Universal Robots PolyScope program: AdientTorsF_Eol1L.urp

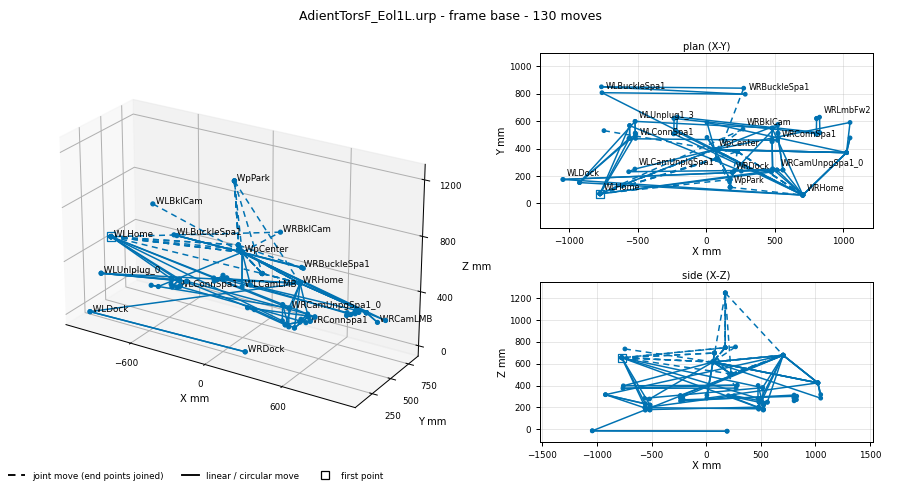
[picture p0: tool path of AdientTorsF_Eol1L.urp in frame base, 130 of 170 moves have a stored position in this frame; points joined in program order, loops and branches not executed]
Program AdientTorsF_Eol1L (installation=EOL_1L directory=/programs createdIn=3.5.1 lastSavedIn=5.26.0 robotSerialNumber=20265101875)
Calibrated DH parameters: a=[-0.000091, -0.609283, -0.566309, 0.000078, -0.000019, 0]; d=[0.180883, 55.684211, -64.380909, 8.871165, 0.119736, 0.115499]; alpha=[1.570556, -0.001038, 0.008646, 1.570192, -1.569654, 0]; deltaTheta=[0, -0.094548, 6.245733, 0.132006, -0.000002, 0]
InitVariablesNode variables(variable(name=Abort, expression=False), variable(name=AdapterReady_L, expression=False), variable(name=AdapterReady_R, expression=False), variable(name=CMD_Heartbt_i1, expression=0), variable(name=CMD_Heartbt_i2, expression=0), variable(name=CMD_Program_i1, expression=0), variable(name=CMD_Program_i2, expression=0), variable(name=CMD_Reserve_i1, expression=0), variable(name=CMD_Reserve_i2, expression=0), variable(name=CMD_Timeout_i1, expression=0), variable(name=CMD_Timeout_i2, expression=0), variable(name=CamCorrectnOK, expression=0), variable(name=DEBUG, expression=False), variable(name=D_rel, expression=p[0,0,0,0,0,0]), variable(name=EvtBeep, expression=False), variable(name=EvtDock, expression=0), variable(name=Mute, expression=False), variable(name=P_ini, expression=get_actual_tcp_pose()), variable(name=Parking, expression=0), variable(name=ProgExe, expression=0), variable(name=STS_Heartbeat, expression=False), variable(name=STS_Progress, expression=0), variable(name=STS_Reservation, expression=0), variable(name=SetCameraProg, expression=0))
BeforeStart
  SuppressedNode
    DEBUG := True
  'SW version, to be used to track changes and keep sync of all stations'
  SW_Ver := 1.0
  Folder Scripts [hidden by the author, left out]
  Folder Avoid guidance screen [hidden by the author, left out]
  Call GripperOpen
  GoToHome := True
  Script: socket_open("127.0.0.1",30001)
Robot Program (runOnlyOnce=false)
  Folder Execute Program
    Folder Init
      Wait Condition expression=EvtDock≤0
      Folder Verify adapter ready
        If digital_in[0] or analog_in[3]<(ivGripSensOpen+0.3)
          AdapterReady_L := False
        If digital_in[4] or analog_in[3]<(ivGripSensOpen+0.3)
          AdapterReady_R := False
      Folder Go to home pos automatically
        If GoToHome and  not (AdapterReady_L or AdapterReady_R)
          Wait Sleep waitTime=1
          If InRange(P_Flange[0],-1,-0.2) and InRange(P_Flange[1],-0.5,0.5) and InRange(P_Flange[2],0.3,1)
            If AdapterDocked or DEBUG or (analog_in[3]<(ivGripSensOpen+0.3))
              MoveJ speed 120 deg/s, acceleration 500 deg/s^2 (useActiveTCP=false positionType=JointAngles optimoveEnabled=false optiMoveSpeed=0.3 optiMoveAcceleration=0.09) tcp=t0_Flange; feature=Base
                Waypoint WLHome: TCP in base x=-773.534 y=70.689 z=655.308 mm, rx=3.1416 ry=0 rz=0 rad; joints [187.663, -96.209, -85.791, -88.066, 90.49, -82.232] deg; TCP offset x=0 y=0 z=0 mm, rx=0 ry=0 rz=3.1416 rad
            Else 
              Popup Error (haltProgram=false message=Adapter must be docked inputType=Text)
              Halt
          ElseIf AtCenterPos
            MoveJ speed 120 deg/s, acceleration 500 deg/s^2 (useActiveTCP=true positionType=JointAngles optimoveEnabled=false optiMoveSpeed=0.3 optiMoveAcceleration=0.09) feature=Base
              Waypoint WpCenter: TCP in base x=62.197 y=393.251 z=616.502 mm, rx=-0.0356 ry=3.1413 rz=-0.0001 rad; joints [106.827, -57.183, -119.283, -93.604, 90.531, 15.582] deg
          ElseIf AtParkPos
            MoveJ speed 120 deg/s, acceleration 500 deg/s^2 (useActiveTCP=true positionType=JointAngles optimoveEnabled=false optiMoveSpeed=0.3 optiMoveAcceleration=0.09) feature=Base
              Waypoint WpPark: TCP in base x=175.046 y=118.455 z=1248.983 mm, rx=-2.2111 ry=2.2293 rz=-0.0002 rad; joints [89.999, -90, 0, -180, 90, -90] deg
          ElseIf InRange(P_Flange[0],0.2,1.2) and InRange(P_Flange[1],-0.5,0.5) and InRange(P_Flange[2],0.3,1)
            If AdapterDocked or DEBUG or (analog_in[3]<(ivGripSensOpen+0.3))
              MoveJ speed 120 deg/s, acceleration 500 deg/s^2 (useActiveTCP=true positionType=JointAngles optimoveEnabled=false optiMoveSpeed=0.3 optiMoveAcceleration=0.09) feature=Base
                Waypoint WRHome: TCP in base x=704.968 y=61.356 z=678.212 mm, rx=-2.2214 ry=-2.2214 rz=0 rad; joints [19.143, -89.513, -90.55, -90.002, 90.503, 19.233] deg; TCP offset x=0 y=0 z=0 mm, rx=0 ry=0 rz=3.1416 rad
            Else 
              Popup Error (haltProgram=false message=Adapter must be docked inputType=Text)
              Halt
          Else 
            Popup Error (haltProgram=false message=Illegal position. Adjust arm to open space in front of the backrest, or [Move]->[Home] inputType=Text)
            Halt
        GoToHome := False
      If DEBUG
        'Popup window with program selection'
        ProgExe :=  (valueSource=Operator message=Program number? valueType=Integer)
      If ProgExe>0
        Folder Init
          Mute := False
          Wait Condition expression=not GoToHome
          If In(ProgExe,[11,12,14])
            AdapterReady_R := False
          ElseIf In(ProgExe,[51,52,54])
            AdapterReady_L := False
          Else 
            AdapterReady_L := False
            AdapterReady_R := False
    Folder Programs
      If InRange(ProgExe,1,99)
        Folder Undock
          If In(ProgExe,[11,51])
            Script: Report(1)
            Folder AtHome?
              Timer (action=Reset) variable(name=T_Timeout)
              Timer (action=Start) variable=T_Timeout
              Wait Condition expression=AtHomePos or T_Timeout>5
              If not AtHomePos
                Script: Report(90)
            If Progress_run() and  not AdapterDocked
              Script: Report(94)
            If Progress_run()
              Folder Undock
                MoveL speed 1000 mm/s, acceleration 3000 mm/s^2 (useActiveTCP=false optimoveEnabled=false optiMoveSpeed=0.3 optiMoveAcceleration=0.09) tcp=t2_Gripper; feature=Base
                  Call GripperOpenQuick
                  If False
                    Waypoint WLDock: TCP in base x=-1043.478 y=175.197 z=-14.02 mm, rx=1.8607 ry=1.8607 rz=0.6057 rad; joints [179.892, -126.837, -85.911, -93.381, 90.434, -0.034] deg; TCP offset x=0 y=-260 z=74 mm, rx=0 ry=0 rz=0 rad
                    Waypoint WRDock: TCP in base x=191.182 y=225.632 z=-17.704 mm, rx=1.8937 ry=1.8608 rz=0.5985 rad; joints [64.532, -92.299, -158.794, -2.395, 58.985, 241.468] deg
                  If ProgExe<50
                    WpDock := WLDock
                    WpHome := WLHome
                  Else 
                    WpDock := WRDock
                    WpHome := WRHome
                  Wp := pose_trans(WpDock, p[0,0.175,-0.1,0,0,0])
                  Waypoint Variable (Variable): motionParameters(blendRadius=0.05); variable=Wp
                  Call GripperOpen
                  Wp := pose_trans(WpDock, p[0,0.075,0.01,0,0,0])
                  Waypoint Variable (Variable): motionParameters(blendRadius=0.01); variable=Wp
                  Wp := pose_trans(WpDock, p[0,0.055,0,0,0,0])
                  Waypoint Variable (Variable): motionParameters(blendRadius=0.01); variable=Wp
                  Waypoint Variable (Variable): variable=WpDock
                  Call GripperClose
                  Wp := pose_trans(WpDock, p[0,0.25,0,0,0,0])
                  Waypoint Variable (Variable): variable=Wp
                If ProgExe<50
                  AdapterReady_L := True
                Else 
                  AdapterReady_R := True
                Script: Report(50)
            Script: Report(50)
        Folder Connect
          If In(ProgExe,[12,14,52,54])
            Script: Report(1)
            If ProgExe<50 and AdapterReady_L
              Undock := False
            ElseIf ProgExe≥50 and AdapterReady_R
              Undock := False
            Else 
              Undock := True
              Folder AtHome? [hidden by the author, left out]
              If Progress_run() and  not AdapterDocked
                Script: Report(94)
            If Progress_run()
              Folder Undock
                If Undock
                  MoveL speed 1000 mm/s, acceleration 3000 mm/s^2 (useActiveTCP=false optimoveEnabled=false optiMoveSpeed=0.3 optiMoveAcceleration=0.09) tcp=t2_Gripper; feature=Base
                    Call GripperOpenQuick
                    If False
                      Waypoint WLDock: TCP in base x=-1043.478 y=175.197 z=-14.02 mm, rx=1.8607 ry=1.8607 rz=0.6057 rad; joints [179.892, -126.837, -85.911, -93.381, 90.434, -0.034] deg; TCP offset x=0 y=-260 z=74 mm, rx=0 ry=0 rz=0 rad
                      Waypoint WRDock: TCP in base x=191.182 y=225.632 z=-17.704 mm, rx=1.8937 ry=1.8608 rz=0.5985 rad; joints [64.532, -92.299, -158.794, -2.395, 58.985, 241.468] deg
                    If ProgExe<50
                      WpDock := WLDock
                      WpHome := WLHome
                    Else 
                      WpDock := WRDock
                      WpHome := WRHome
                    Wp := pose_trans(WpDock, p[0,0.175,-0.1,0,0,0])
                    Waypoint Variable (Variable): motionParameters(blendRadius=0.05); variable=Wp
                    Call GripperOpen
                    Wp := pose_trans(WpDock, p[0,0.075,0.01,0,0,0])
                    Waypoint Variable (Variable): motionParameters(blendRadius=0.01); variable=Wp
                    Wp := pose_trans(WpDock, p[0,0.055,0,0,0,0])
                    Waypoint Variable (Variable): motionParameters(blendRadius=0.01); variable=Wp
                    Waypoint Variable (Variable): variable=WpDock
                    Call GripperClose
                    Wp := pose_trans(WpDock, p[0,0.25,0,0,0,0])
                    Waypoint Variable (Variable): variable=Wp
                AdapterReady_L := False
                AdapterReady_R := False
                Script: Report(2)
              CamCorrection := p[0,0,0,0,0,0]
              SuppressedNode
                Folder Camera
                  MoveL speed 250 mm/s, acceleration 1200 mm/s^2 (useActiveTCP=false optimoveEnabled=false optiMoveSpeed=0.3 optiMoveAcceleration=0.09) tcp=t0_Flange; feature=Base
                    If In(ProgExe,[12,13])
                      SetCameraProg := 12
                      Waypoint WLCamConSpa1: TCP in base x=-511.083 y=256.44 z=253.227 mm, rx=2.1948 ry=2.1949 rz=-0.0574 rad; joints [170.312, -93.988, -133.728, -42.837, 93.248, -9.279] deg; TCP offset x=0 y=0 z=0 mm, rx=0 ry=0 rz=0 rad
                    If In(ProgExe,[14])
                      SetCameraProg := ProgExe
                      Waypoint WLCamConSpa3: TCP in base x=-559.049 y=229.366 z=263.196 mm, rx=-2.2214 ry=-2.2215 rz=0 rad; joints [174.302, -95.829, -130.307, -43.928, 90.296, -5.276] deg
                    If In(ProgExe,[52,53])
                      SetCameraProg := 52
                      Waypoint WRCamConSpa1: TCP in base x=528.577 y=256.538 z=254.589 mm, rx=2.1946 ry=2.1948 rz=-0.0575 rad; joints [43.439, -94.974, -131.929, -45.242, 88.117, 223.892] deg
                    If In(ProgExe,[54])
                      SetCameraProg := ProgExe
                      Waypoint WRCamConSpa3: TCP in base x=480.455 y=221.374 z=266.967 mm, rx=-2.2214 ry=-2.2215 rz=-0.0001 rad; joints [43.801, -88.335, -137.68, -44.047, 90.305, 224.222] deg
                  Call CamAcquire
                  CamCorrection := p[CamData[0],CamData[1]*-0.5,CamData[1],0,0,0]
            SuppressedNode
              If Progress_run() and CamCorrectnOK≠ProgExe
                EvtDock := 1
                Wait Condition expression=EvtDock≟0
                Script: Report(91)
            Folder Connect
              If Progress_run()
                Set NoAction tcp=t2_Gripper
                MoveL speed 1000 mm/s, acceleration 3000 mm/s^2 (useActiveTCP=false optimoveEnabled=false optiMoveSpeed=0.3 optiMoveAcceleration=0.09) tcp=t2_Gripper; feature=Base
                  If False
                    'wp is set to position exactly 30mm below'
                    Waypoint WLConnSpa1: motionParameters(blendRadius=0.045); TCP in base x=-514.347 y=474.559 z=185.987 mm, rx=3.0892 ry=0 rz=0.0001 rad; joints [174.313, -90.885, -134.162, -45.296, 93.296, -95.282] deg; TCP offset x=0 y=260 z=74 mm, rx=0 ry=0 rz=3.1416 rad
                    Waypoint WLConnSpa3: TCP in base x=-563.167 y=472.162 z=197.967 mm, rx=2.9544 ry=0 rz=0.0002 rad; joints [172.16, -92.445, -126.338, -52.702, 100.982, -97.611] deg
                    Waypoint WRConnSpa1: TCP in base x=520.916 y=460.286 z=187.058 mm, rx=3.089 ry=0 rz=-0.0005 rad; joints [39.919, -90.524, -133.875, -47.63, 88.028, 130.365] deg
                    Waypoint WRConnSpa3: TCP in base x=478.559 y=467.416 z=198.199 mm, rx=3.0125 ry=0.0525 rz=-0.0035 rad; joints [44.279, -85.291, -133.969, -56.002, 85.12, 132.879] deg
                  If In(ProgExe,[12])
                    Wp := pose_trans(WLConnSpa1, CamCorrection)
                  If In(ProgExe,[14])
                    Wp := pose_add(WLConnSpa3, CamCorrection)
                  If In(ProgExe,[52])
                    Wp := pose_trans(WRConnSpa1, CamCorrection)
                  If In(ProgExe,[54])
                    Wp := pose_add(WRConnSpa3, CamCorrection)
                  Waypoint Variable (Variable): variable=Wp
                Force Frame feature=Joint_6_name; selection=[0, 0, 1, 0, 0, 0]; wrench=[0, 0, -30, 0, 0, 0]; limitsForce=[0.15, 0.15, 0.1, 1.047198, 1.047198, 1.047198]; limitsMotion=[0.1, 0.1, 0.1, 0.349066, 0.349066, 0.349066]
                  Wait Sleep waitTime=1
                Force Frame feature=Joint_6_name; selection=[1, 0, 1, 0, 0, 0]; wrench=[0, 0, -30, 0, 0, 0]; limitsForce=[0.15, 0.15, 0.05, 1.047198, 1.047198, 1.047198]; limitsMotion=[0.1, 0.1, 0.1, 0.349066, 0.349066, 0.349066]
                  Wait Sleep waitTime=0.5
                'position ok'
                If InRange(Wp[2]+0.03-P_act[2],-0.015,0.015)
                  'ok'
                Else 
                  EvtDock := 2
                  Wait Condition expression=EvtDock≤0
                  Script: Report(96)
              If Progress_run()
                Force Frame feature=Joint_6_name; selection=[0, 1, 0, 0, 0, 0]; wrench=[0, -60, -10, 0, 0, 0]; limitsForce=[0.15, 0.05, 0.01, 1.047198, 1.047198, 1.047198]; limitsMotion=[0.1, 0.1, 0.1, 0.349066, 0.349066, 0.349066]
                  Wait Sleep waitTime=1
                MoveL speed 1000 mm/s, acceleration 3000 mm/s^2 (useActiveTCP=true optimoveEnabled=false optiMoveSpeed=0.3 optiMoveAcceleration=0.09) feature=Base
                  Wp := pose_trans(P_act, p[0,0.005,0,0,0,0])
                  Waypoint Variable (Variable): variable=Wp
                Call GripperOpen
                Force Frame feature=Joint_6_name; selection=[0, 1, 0, 0, 0, 0]; wrench=[0, -60, -10, 0, 0, 0]; limitsForce=[0.15, 0.1, 0.01, 1.047198, 1.047198, 1.047198]; limitsMotion=[0.1, 0.1, 0.1, 0.349066, 0.349066, 0.349066]
                  Wait Sleep waitTime=1
                  Script: Report(5)
                  MoveL speed 500 mm/s, acceleration 2000 mm/s^2 (useActiveTCP=true optimoveEnabled=false optiMoveSpeed=0.3 optiMoveAcceleration=0.09) feature=Base
                    Wp0 := get_actual_tcp_pose()
                    Wp := pose_trans(Wp0, p[0,0,0,0,0,0.07])
                    Waypoint Variable (Variable): variable=Wp
                    Wp := pose_trans(Wp0, p[0,0,0,0,0,-0.07])
                    Waypoint Variable (Variable): variable=Wp
                    Waypoint Variable (Variable): variable=Wp0
                    Wp := pose_trans(Wp0, p[0,0,0.01,0,0,0])
                    Waypoint Variable (Variable): variable=Wp
                    Waypoint Variable (Variable): variable=Wp0
                MoveL speed 1000 mm/s, acceleration 3000 mm/s^2 (useActiveTCP=true optimoveEnabled=false optiMoveSpeed=0.3 optiMoveAcceleration=0.09) feature=Base
                  Wp0 := get_actual_tcp_pose()
                  Wp := pose_trans(Wp0, p[0,0.015,0,0,0,0])
                  Waypoint Variable (Variable): variable=Wp
                Force Frame feature=Joint_6_name; selection=[0, 1, 0, 0, 0, 0]; wrench=[0, -60, 0, 0, 0, 0]; limitsForce=[0.15, 0.5, 0.15, 1.047198, 1.047198, 1.047198]; limitsMotion=[0.1, 0.1, 0.1, 0.349066, 0.349066, 0.349066]
                  Wait Sleep waitTime=0.5
                Script: Report(6)
                Timer (action=Reset) variable=T_Timeout
                Timer (action=Start) variable=T_Timeout
                Folder Test switch pin, retreat on fail
                  Wait Condition expression=Flags[0] or T_Timeout>10 or DEBUG
                  If not Flags[0] and  not DEBUG
                    EvtDock := 2
                    Wait Condition expression=EvtDock≤0
                    Script: Report(95)
            If Progress_run()
              MoveL speed 1000 mm/s, acceleration 3000 mm/s^2 (useActiveTCP=false optimoveEnabled=false optiMoveSpeed=0.3 optiMoveAcceleration=0.09) tcp=t0_Flange; feature=Base
                Set NoAction tcp=t0_Flange
                P_act := get_actual_tcp_pose()
                Wp := pose_trans(P_act, p[0,0.1,0,0,0,0])
                Waypoint Variable (Variable): motionParameters(blendRadius=0.05); variable=Wp
                Wp := pose_trans(Wp, p[0,0.1,-0.1,0,0,0])
                Waypoint Variable (Variable): motionParameters(blendRadius=0.05); variable=Wp
                Waypoint Variable (Variable): variable=WpHome
              Script: Report(50)
        Folder Buckle
          If In(ProgExe,[15,16,55,56])
            Script: Report(1)
            Folder AtHome?
              Timer (action=Reset) variable=T_Timeout
              Timer (action=Start) variable=T_Timeout
              Wait Condition expression=AtHomePos or (In(ProgExe,[55,56]) and AtCenterPos) or T_Timeout>5
              If AtHomePos or (In(ProgExe,[55,56]) and AtCenterPos)
                'nop'
              Else 
                Script: Report(90)
            If Progress_run() and  not ((digital_in[2] and ProgExe<50)  or (digital_in[6] and ProgExe>50))
              Script: Report(92)
            If Progress_run()
              Call GripperCloseQuick
              Folder Camera
                SetCameraProg := ProgExe
                MoveL speed 1000 mm/s, acceleration 3000 mm/s^2 (useActiveTCP=false optimoveEnabled=false optiMoveSpeed=0.3 optiMoveAcceleration=0.09) tcp=t0_Flange; feature=Base
                  If ProgExe<50
                    Waypoint WLBklCam: TCP in base x=-744.742 y=530.901 z=735.863 mm, rx=-1.8029 ry=-0.697 rz=1.8635 rad; joints [151.622, -114.453, -78.198, 13.926, 120.764, -128.64] deg; TCP offset x=0 y=0 z=0 mm, rx=0 ry=0 rz=3.1416 rad
                  Else 
                    MoveJ speed 120 deg/s, acceleration 500 deg/s^2 (useActiveTCP=false positionType=JointAngles optimoveEnabled=false optiMoveSpeed=0.3 optiMoveAcceleration=0.09) tcp=t0_Flange; feature=Base
                      Waypoint WpCenter: motionParameters(blendRadius=0.1); TCP in base x=62.197 y=393.251 z=616.502 mm, rx=-0.0356 ry=3.1413 rz=-0.0001 rad; joints [106.827, -57.183, -119.283, -93.604, 90.531, 15.582] deg
                      Waypoint WRBklCam: motionParameters(jointSpeed=3.141593 jointAcceleration=17.453293 cartesianSpeed=0.25 cartesianAcceleration=1.2); TCP in base x=268.762 y=542.285 z=754.984 mm, rx=0.5116 ry=1.5528 rz=0.4744 rad; joints [92.2, -78.985, -94.967, -140.229, 4.149, 80.102] deg
                Call GripperClose
                Call CamAcquire
                Call CamCalculateCorectnPlane
              If CamCorrectnOK≟ProgExe and InRange(CamCorrection[1],-0.05,0.05) and InRange(CamCorrection[2],-0.03,0.03)
                'empty'
              Else 
                CamCorrectnOK := 0
                MoveJ speed 120 deg/s, acceleration 500 deg/s^2 (useActiveTCP=false positionType=JointAngles optimoveEnabled=false optiMoveSpeed=0.3 optiMoveAcceleration=0.09) tcp=t0_Flange; feature=Base
                  If ProgExe<50
                    Waypoint WLHome: TCP in base x=-773.534 y=70.689 z=655.308 mm, rx=3.1416 ry=0 rz=0 rad; joints [187.663, -96.209, -85.791, -88.066, 90.49, -82.232] deg
                  Else 
                    Waypoint WRBklMidp3: TCP in base x=75.853 y=323.344 z=698.705 mm, rx=3.1416 ry=0 rz=0 rad; joints [108.301, -50.923, -113.164, -105.98, 90.537, -161.757] deg
                    Waypoint WpCenter: motionParameters(jointSpeed=3.141593 jointAcceleration=17.453293 cartesianSpeed=0.25 cartesianAcceleration=1.2); TCP in base x=62.197 y=393.251 z=616.502 mm, rx=-0.0356 ry=3.1413 rz=-0.0001 rad; joints [106.827, -57.183, -119.283, -93.604, 90.531, 15.582] deg
                    STS_Reservation := 0
                Script: Report(91)
              If CamCorrectnOK≟ProgExe
                Folder Insert
                  MoveL speed 1000 mm/s, acceleration 3000 mm/s^2 (useActiveTCP=false optimoveEnabled=false optiMoveSpeed=0.3 optiMoveAcceleration=0.09) tcp=t3_Blade; feature=Base
                    If False
                      'must be set with blade ca one half into buckle slot'
                      Waypoint WLBuckleSpa1: TCP in base x=-759.148 y=807.506 z=398.072 mm, rx=-2.6459 ry=0.0002 rz=0.0002 rad; joints [153.1, -131.84, -57.173, -67.423, 65.296, -119.666] deg; TCP offset x=-134 y=56 z=118 mm, rx=0 ry=0 rz=3.1416 rad
                      Waypoint WRBuckleSpa1: TCP in base x=285.068 y=796.337 z=403.859 mm, rx=-2.6293 ry=0.0331 rz=0.1099 rad; joints [90.6, -91.771, -115.486, -33.413, 94.028, -176.49] deg; TCP offset x=-134 y=56 z=118 mm, rx=0 ry=0 rz=3.1416 rad
                      Waypoint WLBuckleSpa3: TCP in base x=-763.082 y=850.426 z=375.25 mm, rx=-2.5567 ry=0.0462 rz=-0.1173 rad; joints [152.045, -137.406, -51.844, -69.177, 58.56, -118.947] deg
                      Waypoint WRBuckleSpa3: TCP in base x=273.907 y=840.505 z=376.981 mm, rx=-2.5518 ry=0.05 rz=0.0053 rad; joints [93.121, -97.682, -115.538, -23.158, 87.96, -174.79] deg
                    If ProgExe≟15
                      Wp := WLBuckleSpa1
                    If ProgExe≟16
                      Wp := WLBuckleSpa3
                    If ProgExe≟55
                      MoveJ speed 180 deg/s, acceleration 1000 deg/s^2 (useActiveTCP=false positionType=JointAngles optimoveEnabled=false optiMoveSpeed=0.3 optiMoveAcceleration=0.09) tcp=t0_Flange; feature=Base
                        Waypoint WRBklMidp3: TCP in base x=75.853 y=323.344 z=698.705 mm, rx=3.1416 ry=0 rz=0 rad; joints [108.301, -50.923, -113.164, -105.98, 90.537, -161.757] deg; TCP offset x=0 y=0 z=0 mm, rx=0 ry=0 rz=3.1416 rad
                      Wp := WRBuckleSpa1
                    If ProgExe≟56
                      MoveJ speed 180 deg/s, acceleration 1000 deg/s^2 (useActiveTCP=true positionType=JointAngles optimoveEnabled=false optiMoveSpeed=0.3 optiMoveAcceleration=0.09) feature=Base
                        Waypoint WRBklMidp3: TCP in base x=75.853 y=323.344 z=698.705 mm, rx=3.1416 ry=0 rz=0 rad; joints [108.301, -50.923, -113.164, -105.98, 90.537, -161.757] deg; TCP offset x=0 y=0 z=0 mm, rx=0 ry=0 rz=3.1416 rad
                      Wp := WRBuckleSpa3
                    Wp0 := pose_trans(Wp,p[0,0,-0.02,0,0,0])
                    Wp0 := pose_add(Wp0,Base_w_correctn)
                    Waypoint Variable (Variable): variable=Wp0
                  Script: Report(5)
                  Timer (action=Reset) variable=T_Timeout
                  Timer (action=Start) variable=T_Timeout
                  Wait Condition expression=Flags[8] or Abort or DEBUG or T_Timeout>25
                  If Flags[8] or DEBUG
                    Script: Report(6)
                    Set NoAction tcp=t3_Blade
                    Force Frame feature=Joint_6_name; selection=[0, 0, 1, 0, 0, 0]; wrench=[0, 0, 15, 0, 0, 0]; limitsForce=[0.15, 0.15, 0.15, 1.047198, 1.047198, 1.047198]; limitsMotion=[0.1, 0.1, 0.1, 0.349066, 0.349066, 0.349066]
                      Wait Sleep waitTime=1
                    If not Flags[9] and  not Abort
                      MoveL speed 50 mm/s, acceleration 500 mm/s^2 (useActiveTCP=false optimoveEnabled=false optiMoveSpeed=0.3 optiMoveAcceleration=0.09) tcp=t3_Blade; feature=Base
                        Waypoint Variable (Variable): variable=Wp
                      Force Frame feature=Joint_6_name; selection=[1, 1, 1, 0, 0, 0]; wrench=[0, 0, 50, 0, 0, 0]; limitsForce=[0.15, 0.15, 0.25, 1.047198, 1.047198, 1.047198]; limitsMotion=[0.1, 0.1, 0.1, 0.349066, 0.349066, 0.349066]
                        Wait Sleep waitTime=1.5
                    If not Flags[9] and  not Abort
                      MoveL speed 50 mm/s, acceleration 500 mm/s^2 (useActiveTCP=false optimoveEnabled=false optiMoveSpeed=0.3 optiMoveAcceleration=0.09) tcp=t3_Blade; feature=Base
                        Waypoint Variable (Variable): variable=Wp
                      Force Frame feature=Joint_6_name; selection=[1, 1, 1, 0, 0, 0]; wrench=[0, 0, 50, 0, 0, 0]; limitsForce=[0.15, 0.15, 0.25, 1.047198, 1.047198, 1.047198]; limitsMotion=[0.1, 0.1, 0.1, 0.349066, 0.349066, 0.349066]
                        Wait Sleep waitTime=1.5
                    If not Flags[9] and  not Abort
                      MoveL speed 50 mm/s, acceleration 500 mm/s^2 (useActiveTCP=false optimoveEnabled=false optiMoveSpeed=0.3 optiMoveAcceleration=0.09) tcp=t3_Blade; feature=Base
                        Waypoint Variable (Variable): variable=Wp
                      Force Frame feature=Joint_6_name; selection=[1, 1, 1, 0, 0, 0]; wrench=[0, 0, 50, 0, 0, 0]; limitsForce=[0.15, 0.15, 0.25, 1.047198, 1.047198, 1.047198]; limitsMotion=[0.1, 0.1, 0.1, 0.349066, 0.349066, 0.349066]
                        Wait Sleep waitTime=1.5
                  MoveL speed 1000 mm/s, acceleration 3000 mm/s^2 (useActiveTCP=false optimoveEnabled=false optiMoveSpeed=0.3 optiMoveAcceleration=0.09) tcp=t3_Blade; feature=Base
                    Waypoint Variable (Variable): variable=Wp
                    MoveDirectionNode (selectedDirection=ZMinus) feature=Joint_6_name
                      Until DISTANCE (allowActions=false deceleration=3 distanceNodeType=STOP) Distance=0.02; motionParameters(blendRadius=0)
                    If In(ProgExe,[15,16])
                      MoveJ speed 120 deg/s, acceleration 500 deg/s^2 (useActiveTCP=false positionType=JointAngles optimoveEnabled=false optiMoveSpeed=0.3 optiMoveAcceleration=0.09) tcp=t0_Flange; feature=Base
                        Waypoint WLHome: TCP in base x=-773.534 y=70.689 z=655.308 mm, rx=3.1416 ry=0 rz=0 rad; joints [187.663, -96.209, -85.791, -88.066, 90.49, -82.232] deg; TCP offset x=0 y=0 z=0 mm, rx=0 ry=0 rz=3.1416 rad
                    If In(ProgExe,[55,56])
                      MoveJ speed 180 deg/s, acceleration 1000 deg/s^2 (useActiveTCP=false positionType=JointAngles optimoveEnabled=false optiMoveSpeed=0.3 optiMoveAcceleration=0.09) tcp=t0_Flange; feature=Base
                        Waypoint WRBklMidp3: TCP in base x=75.853 y=323.344 z=698.705 mm, rx=3.1416 ry=0 rz=0 rad; joints [108.301, -50.923, -113.164, -105.98, 90.537, -161.757] deg
                        Waypoint WpCenter: TCP in base x=62.197 y=393.251 z=616.502 mm, rx=-0.0356 ry=3.1413 rz=-0.0001 rad; joints [106.827, -57.183, -119.283, -93.604, 90.531, 15.582] deg
                        STS_Reservation := 0
                  If Progress_check()≥6
                    Script: Report(50)
                  Else 
                    Script: Report(95)
        Folder Disconnect
          If In(ProgExe,[21,22,23,61,62,63])
            Script: Report(1)
            Folder AtHome? [hidden by the author, left out]
            If Progress_run()
              If In(ProgExe,[21,22])
                SetCameraProg := 21
                MoveL speed 1000 mm/s, acceleration 3000 mm/s^2 (useActiveTCP=false optimoveEnabled=false optiMoveSpeed=0.3 optiMoveAcceleration=0.09) tcp=t0_Flange; feature=Base
                  Waypoint WLCamUnplgSpa1: TCP in base x=-519.312 y=251.237 z=277.522 mm, rx=2.1002 ry=2.1002 rz=-0.2414 rad; joints [168.952, -92.992, -131.142, -48.398, 103.196, -10.943] deg
              If In(ProgExe,[23])
                SetCameraProg := ProgExe
                MoveL speed 1000 mm/s, acceleration 3000 mm/s^2 (useActiveTCP=false optimoveEnabled=false optiMoveSpeed=0.3 optiMoveAcceleration=0.09) tcp=t0_Flange; feature=Base
                  SuppressedNode
                    Waypoint WLCamUnpgSpa3_0: motionParameters(blendRadius=0.05); TCP in base x=-374.135 y=332.475 z=451.177 mm, rx=2.1642 ry=2.1642 rz=-0.1205 rad; joints [157.169, -73.07, -127.046, -72.385, 96.229, -22.692] deg
                  Waypoint WLCamUnpgSpa3: TCP in base x=-564.455 y=231.557 z=283.493 mm, rx=2.1235 ry=2.1236 rz=-0.1987 rad; joints [172.076, -95.315, -127.907, -48.261, 100.917, -7.669] deg
              If In(ProgExe,[61,62])
                SetCameraProg := 61
                MoveL speed 1000 mm/s, acceleration 3000 mm/s^2 (useActiveTCP=false optimoveEnabled=false optiMoveSpeed=0.3 optiMoveAcceleration=0.09) tcp=t0_Flange; feature=Base
                  Waypoint WRCamUnpgSpa1_0: motionParameters(blendRadius=0.05); TCP in base x=516.477 y=243.64 z=380.929 mm, rx=2.1642 ry=2.1642 rz=-0.1204 rad; joints [43.859, -83.9, -126.098, -64.514, 85.844, 224.336] deg
                  Waypoint WRCamUnplgSpa1: TCP in base x=516.477 y=243.64 z=244.776 mm, rx=2.1642 ry=2.1642 rz=-0.1204 rad; joints [43.842, -94.277, -133.514, -46.729, 85.729, 224.433] deg
              If In(ProgExe,[63])
                SetCameraProg := ProgExe
                MoveL speed 1000 mm/s, acceleration 3000 mm/s^2 (useActiveTCP=false optimoveEnabled=false optiMoveSpeed=0.3 optiMoveAcceleration=0.09) tcp=t0_Flange; feature=Base
                  Waypoint WRCamUnpgSpa3_0: motionParameters(blendRadius=0.05); TCP in base x=475.545 y=231.557 z=401.094 mm, rx=2.1235 ry=2.1236 rz=-0.1987 rad; joints [46.754, -78.431, -127.605, -71.891, 83.171, 227.5] deg
                  Waypoint WRCamUnpgSpa3: TCP in base x=475.545 y=229.337 z=283.493 mm, rx=2.1235 ry=2.1236 rz=-0.1987 rad; joints [46.564, -86.446, -135.161, -56.311, 83.062, 227.425] deg
              Call CamAcquire
              Call CamCalculateCorectnPlane
            If Progress_run() and CamCorrectnOK≠ProgExe
              MoveL speed 1000 mm/s, acceleration 3000 mm/s^2 (useActiveTCP=false optimoveEnabled=false optiMoveSpeed=0.3 optiMoveAcceleration=0.09) tcp=t0_Flange; feature=Base
                If ProgExe<50
                  Waypoint WLHome: TCP in base x=-773.534 y=70.689 z=655.308 mm, rx=3.1416 ry=0 rz=0 rad; joints [187.663, -96.209, -85.791, -88.066, 90.49, -82.232] deg; TCP offset x=0 y=0 z=0 mm, rx=0 ry=0 rz=3.1416 rad
                Else 
                  MoveL speed 1000 mm/s, acceleration 3000 mm/s^2 (useActiveTCP=false optimoveEnabled=false optiMoveSpeed=0.3 optiMoveAcceleration=0.09) tcp=t0_Flange; feature=Base
                    Waypoint WRCamUnpgSpa1_0: motionParameters(blendRadius=0.05); TCP in base x=516.477 y=243.64 z=380.929 mm, rx=2.1642 ry=2.1642 rz=-0.1204 rad; joints [43.859, -83.9, -126.098, -64.514, 85.844, 224.336] deg
                  Waypoint WRHome: TCP in base x=704.968 y=61.356 z=678.212 mm, rx=-2.2214 ry=-2.2214 rz=0 rad; joints [19.143, -89.513, -90.55, -90.002, 90.503, 19.233] deg; TCP offset x=0 y=0 z=0 mm, rx=0 ry=0 rz=3.1416 rad
              Script: Report(91)
            If Progress_run()
              Call GripperOpenQuick
              Folder Disconnect
                If In(ProgExe,[21,22])
                  MoveL speed 1000 mm/s, acceleration 3000 mm/s^2 (useActiveTCP=false optimoveEnabled=false optiMoveSpeed=0.3 optiMoveAcceleration=0.09) tcp=t2_Gripper; feature=Base_w_correctn
                    Waypoint WLUnlplug_0: motionParameters(blendRadius=0.05); TCP in base x=-922.864 y=152.307 z=316.977 mm, rx=2.2214 ry=2.2214 rz=0 rad; joints [181.781, -93.99, -116.062, -60.013, 90.397, 2.107] deg; TCP offset x=0 y=-260 z=74 mm, rx=0 ry=0 rz=0 rad
                    Call GripperOpen
                    Waypoint WLUnplug1_1: motionParameters(blendRadius=0.03); TCP in base x=-515.238 y=504.129 z=221.991 mm, rx=2.6768 ry=0 rz=-0.0006 rad; joints [161.335, -87.939, -119.929, -71.208, 115.593, -110.465] deg; TCP offset x=0 y=260 z=74 mm, rx=0 ry=0 rz=3.1416 rad
                    Waypoint WLUnplug1_2: motionParameters(blendRadius=0.015); TCP in base x=-516.569 y=512.274 z=177.183 mm, rx=2.6768 ry=0 rz=0 rad; joints [160.643, -90.949, -122.086, -66.343, 115.459, 68.823] deg; TCP offset x=0 y=-260 z=74 mm, rx=0 ry=0 rz=0 rad
                    Waypoint WLUnplug1_3: TCP in base x=-517.731 y=598.443 z=180.678 mm, rx=3.0593 ry=-0.0005 rz=0.0001 rad; joints [161.547, -96.621, -127.223, -47.688, 94.795, 71.907] deg
                If In(ProgExe,[23])
                  MoveL speed 1000 mm/s, acceleration 3000 mm/s^2 (useActiveTCP=false optimoveEnabled=false optiMoveSpeed=0.3 optiMoveAcceleration=0.09) tcp=t2_Gripper; feature=Base_w_correctn
                    Waypoint WLUnlplug_0: motionParameters(blendRadius=0.05); TCP in base x=-922.864 y=152.307 z=316.977 mm, rx=2.2214 ry=2.2214 rz=0 rad; joints [181.781, -93.99, -116.062, -60.013, 90.397, 2.107] deg
                    Call GripperOpen
                    Waypoint WLUnplg3_1: motionParameters(blendRadius=0.05); TCP in base x=-558.094 y=476.014 z=233.764 mm, rx=2.6768 ry=0 rz=0 rad; joints [165.009, -89.56, -117.426, -70.357, 116.114, 73.568] deg
                    Waypoint WLUnplg3_2: motionParameters(blendRadius=0.005); TCP in base x=-557.642 y=476.233 z=176.69 mm, rx=2.6768 ry=0 rz=0 rad; joints [164.972, -92.601, -120.933, -63.804, 116.077, 73.582] deg
                    Waypoint WLUnplg3_3: TCP in base x=-557.64 y=567.874 z=198.677 mm, rx=2.9513 ry=0 rz=0 rad; joints [163.24, -95.853, -121.965, -55.361, 100.806, -106.7] deg; TCP offset x=0 y=260 z=74 mm, rx=0 ry=0 rz=3.1416 rad
                If In(ProgExe,[61,62])
                  MoveL speed 1000 mm/s, acceleration 3000 mm/s^2 (useActiveTCP=false optimoveEnabled=false optiMoveSpeed=0.3 optiMoveAcceleration=0.09) tcp=t2_Gripper; feature=Base_w_correctn
                    Waypoint WRUnpgSpa1_0: motionParameters(blendRadius=0.05); TCP in base x=256.479 y=235.425 z=307.381 mm, rx=2.1642 ry=2.1642 rz=-0.1204 rad; joints [43.859, -83.9, -126.098, -64.514, 85.844, 224.336] deg; TCP offset x=0 y=-260 z=74 mm, rx=0 ry=0 rz=0 rad
                    Call GripperOpen
                    Waypoint WRUnpgSpa1_1: motionParameters(blendRadius=0.05); TCP in base x=559.86 y=244.266 z=247.805 mm, rx=1.9727 ry=1.054 rz=0.549 rad; joints [40.557, -86.579, -121.116, -41.845, 38.217, 64.714] deg; TCP offset x=0 y=260 z=74 mm, rx=0 ry=0 rz=3.1416 rad
                    Waypoint WRUnpgSpa1_2: motionParameters(blendRadius=0.03); TCP in base x=524.815 y=481.473 z=221.99 mm, rx=2.6768 ry=0 rz=0 rad; joints [48.645, -86.963, -118.221, -85.548, 73.288, 321.949] deg; TCP offset x=0 y=-260 z=74 mm, rx=0 ry=0 rz=0 rad
                    Waypoint WRUnpgSpa1_3: motionParameters(blendRadius=0.02); TCP in base x=523.431 y=512.274 z=177.183 mm, rx=2.6768 ry=0 rz=0 rad; joints [50.625, -90.73, -119.487, -81.085, 73.982, 323.92] deg; TCP offset x=0 y=-260 z=74 mm, rx=0 ry=0 rz=0 rad
                    Waypoint WRUnpgSpa1_4: TCP in base x=523.021 y=574.6 z=182.646 mm, rx=3.0593 ry=-0.0005 rz=0.0001 rad; joints [48.549, -95.333, -127.836, -50.454, 87.221, 319.057] deg; TCP offset x=0 y=-260 z=74 mm, rx=0 ry=0 rz=0 rad
                If In(ProgExe,[63])
                  MoveL speed 1000 mm/s, acceleration 3000 mm/s^2 (useActiveTCP=false optimoveEnabled=false optiMoveSpeed=0.3 optiMoveAcceleration=0.09) tcp=t2_Gripper; feature=Base_w_correctn
                    Waypoint WRUnpg3_0: motionParameters(blendRadius=0.05); TCP in base x=203.178 y=235.425 z=307.381 mm, rx=2.1642 ry=2.1642 rz=-0.1204 rad; joints [48.044, -78.714, -130.246, -65.872, 86.191, 228.509] deg
                    Call GripperOpen
                    Waypoint WRUnpg3_1: motionParameters(blendRadius=0.05); TCP in base x=484.471 y=251.759 z=247.938 mm, rx=1.9943 ry=1.0212 rz=0.5679 rad; joints [46.405, -77.678, -126.927, -52.297, 36.548, 255.917] deg
                    Waypoint WRUnpg3_2: TCP in base x=480.585 y=451.056 z=185.786 mm, rx=2.6768 ry=0 rz=0 rad; joints [50.025, -83.245, -125.54, -82.347, 73.777, 323.323] deg
                    Waypoint WRUnpg3_4: TCP in base x=480.582 y=549.49 z=202.644 mm, rx=2.9643 ry=0 rz=0 rad; joints [51.538, -87.895, -128.855, -61.335, 84.121, 322.301] deg
                Script: Report(20)
                Wait Condition expression=Flags[7] or DEBUG
              EvtDock := 2
              Wait Condition expression=EvtDock≤0
              If EvtDock<0
                If In(ProgExe,[21,22])
                  MoveL speed 1000 mm/s, acceleration 3000 mm/s^2 (useActiveTCP=false optimoveEnabled=false optiMoveSpeed=0.3 optiMoveAcceleration=0.09) tcp=t2_Gripper; feature=Base_w_correctn
                    Waypoint WLUnplug1_3: TCP in base x=-517.731 y=598.443 z=180.678 mm, rx=3.0593 ry=-0.0005 rz=0.0001 rad; joints [161.547, -96.621, -127.223, -47.688, 94.795, 71.907] deg
                    Waypoint WLUnplug1_2: motionParameters(blendRadius=0); TCP in base x=-516.569 y=512.274 z=177.183 mm, rx=2.6768 ry=0 rz=0 rad; joints [160.643, -90.949, -122.086, -66.343, 115.459, 68.823] deg
                    Waypoint WLUnplug1_1: TCP in base x=-515.238 y=504.129 z=221.991 mm, rx=2.6768 ry=0 rz=-0.0006 rad; joints [161.335, -87.939, -119.929, -71.208, 115.593, -110.465] deg; TCP offset x=0 y=260 z=74 mm, rx=0 ry=0 rz=3.1416 rad
                    SuppressedNode
                      Waypoint WLUnlplug_0: TCP in base x=-922.864 y=152.307 z=316.977 mm, rx=2.2214 ry=2.2214 rz=0 rad; joints [181.781, -93.99, -116.062, -60.013, 90.397, 2.107] deg; TCP offset x=0 y=-260 z=74 mm, rx=0 ry=0 rz=0 rad
                  MoveL speed 1000 mm/s, acceleration 3000 mm/s^2 (useActiveTCP=false optimoveEnabled=false optiMoveSpeed=0.3 optiMoveAcceleration=0.09) tcp=t0_Flange; feature=Base
                    Waypoint WLHome referenceName=WLHome: TCP in base x=-773.534 y=70.689 z=655.308 mm, rx=3.1416 ry=0 rz=0 rad; joints [187.663, -96.209, -85.791, -88.066, 90.49, -82.232] deg; TCP offset x=0 y=0 z=0 mm, rx=0 ry=0 rz=3.1416 rad
                If In(ProgExe,[23])
                  MoveL speed 1000 mm/s, acceleration 3000 mm/s^2 (useActiveTCP=false optimoveEnabled=false optiMoveSpeed=0.3 optiMoveAcceleration=0.09) tcp=t2_Gripper; feature=Base_w_correctn
                    Waypoint WLUnplg3_3: TCP in base x=-557.64 y=567.874 z=198.677 mm, rx=2.9513 ry=0 rz=0 rad; joints [163.24, -95.853, -121.965, -55.361, 100.806, -106.7] deg; TCP offset x=0 y=260 z=74 mm, rx=0 ry=0 rz=3.1416 rad
                    Waypoint WLUnplg3_2: TCP in base x=-557.642 y=476.233 z=176.69 mm, rx=2.6768 ry=0 rz=0 rad; joints [164.972, -92.601, -120.933, -63.804, 116.077, 73.582] deg; TCP offset x=0 y=-260 z=74 mm, rx=0 ry=0 rz=0 rad
                    Waypoint WLUnplg3_1: TCP in base x=-558.094 y=476.014 z=233.764 mm, rx=2.6768 ry=0 rz=0 rad; joints [165.009, -89.56, -117.426, -70.357, 116.114, 73.568] deg
                    SuppressedNode
                      Waypoint WLUnlplug_0: TCP in base x=-922.864 y=152.307 z=316.977 mm, rx=2.2214 ry=2.2214 rz=0 rad; joints [181.781, -93.99, -116.062, -60.013, 90.397, 2.107] deg
                  MoveL speed 1000 mm/s, acceleration 3000 mm/s^2 (useActiveTCP=false optimoveEnabled=false optiMoveSpeed=0.3 optiMoveAcceleration=0.09) tcp=t0_Flange; feature=Base
                    Waypoint WLHome: TCP in base x=-773.534 y=70.689 z=655.308 mm, rx=3.1416 ry=0 rz=0 rad; joints [187.663, -96.209, -85.791, -88.066, 90.49, -82.232] deg; TCP offset x=0 y=0 z=0 mm, rx=0 ry=0 rz=3.1416 rad
                If In(ProgExe,[61,62])
                  MoveL speed 1000 mm/s, acceleration 3000 mm/s^2 (useActiveTCP=false optimoveEnabled=false optiMoveSpeed=0.3 optiMoveAcceleration=0.09) tcp=t2_Gripper; feature=Base_w_correctn
                    Waypoint WRUnpgSpa1_4: TCP in base x=523.021 y=574.6 z=182.646 mm, rx=3.0593 ry=-0.0005 rz=0.0001 rad; joints [48.549, -95.333, -127.836, -50.454, 87.221, 319.057] deg; TCP offset x=0 y=-260 z=74 mm, rx=0 ry=0 rz=0 rad
                    Waypoint WRUnpgSpa1_3: motionParameters(blendRadius=0); TCP in base x=523.431 y=512.274 z=177.183 mm, rx=2.6768 ry=0 rz=0 rad; joints [50.625, -90.73, -119.487, -81.085, 73.982, 323.92] deg; TCP offset x=0 y=-260 z=74 mm, rx=0 ry=0 rz=0 rad
                    Waypoint WRUnpgSpa1_2: motionParameters(blendRadius=0.03); TCP in base x=524.815 y=481.473 z=221.99 mm, rx=2.6768 ry=0 rz=0 rad; joints [48.645, -86.963, -118.221, -85.548, 73.288, 321.949] deg; TCP offset x=0 y=-260 z=74 mm, rx=0 ry=0 rz=0 rad
                    Waypoint WRUnpgSpa1_1: TCP in base x=559.86 y=244.266 z=247.805 mm, rx=1.9727 ry=1.054 rz=0.549 rad; joints [40.557, -86.579, -121.116, -41.845, 38.217, 64.714] deg; TCP offset x=0 y=260 z=74 mm, rx=0 ry=0 rz=3.1416 rad
                    SuppressedNode
                      Waypoint WRUnpgSpa1_0: TCP in base x=256.479 y=235.425 z=307.381 mm, rx=2.1642 ry=2.1642 rz=-0.1204 rad; joints [43.859, -83.9, -126.098, -64.514, 85.844, 224.336] deg; TCP offset x=0 y=-260 z=74 mm, rx=0 ry=0 rz=0 rad
                  MoveL speed 1000 mm/s, acceleration 3000 mm/s^2 (useActiveTCP=false optimoveEnabled=false optiMoveSpeed=0.3 optiMoveAcceleration=0.09) tcp=t0_Flange; feature=Base
                    Waypoint WRHome: TCP in base x=704.968 y=61.356 z=678.212 mm, rx=-2.2214 ry=-2.2214 rz=0 rad; joints [19.143, -89.513, -90.55, -90.002, 90.503, 19.233] deg; TCP offset x=0 y=0 z=0 mm, rx=0 ry=0 rz=3.1416 rad
                If In(ProgExe,[63])
                  MoveL speed 1000 mm/s, acceleration 3000 mm/s^2 (useActiveTCP=false optimoveEnabled=false optiMoveSpeed=0.3 optiMoveAcceleration=0.09) tcp=t2_Gripper; feature=Base_w_correctn
                    Waypoint WRUnpg3_4: TCP in base x=480.582 y=549.49 z=202.644 mm, rx=2.9643 ry=0 rz=0 rad; joints [51.538, -87.895, -128.855, -61.335, 84.121, 322.301] deg; TCP offset x=0 y=-260 z=74 mm, rx=0 ry=0 rz=0 rad
                    Waypoint WRUnpg3_2: TCP in base x=480.585 y=451.056 z=185.786 mm, rx=2.6768 ry=0 rz=0 rad; joints [50.025, -83.245, -125.54, -82.347, 73.777, 323.323] deg
                    Waypoint WRUnpg3_1: TCP in base x=484.471 y=251.759 z=247.938 mm, rx=1.9943 ry=1.0212 rz=0.5679 rad; joints [46.405, -77.678, -126.927, -52.297, 36.548, 255.917] deg
                    SuppressedNode
                      Waypoint WRUnpg3_0: TCP in base x=203.178 y=235.425 z=307.381 mm, rx=2.1642 ry=2.1642 rz=-0.1204 rad; joints [48.044, -78.714, -130.246, -65.872, 86.191, 228.509] deg
                  MoveL speed 1000 mm/s, acceleration 3000 mm/s^2 (useActiveTCP=false optimoveEnabled=false optiMoveSpeed=0.3 optiMoveAcceleration=0.09) tcp=t0_Flange; feature=Base
                    Waypoint WRHome: TCP in base x=704.968 y=61.356 z=678.212 mm, rx=-2.2214 ry=-2.2214 rz=0 rad; joints [19.143, -89.513, -90.55, -90.002, 90.503, 19.233] deg; TCP offset x=0 y=0 z=0 mm, rx=0 ry=0 rz=3.1416 rad
                Script: Report(97)
            If Progress_run()
              Script: Report(50)
        Folder Buttons
          If In(ProgExe,[31,32,37,38,71,72,77,78])
            Script: Report(1)
            Folder AtHome?
              Timer (action=Reset) variable=T_Timeout
              Timer (action=Start) variable=T_Timeout
              Wait Condition expression=AtHomePos or (AtCenterPos and In(ProgExe,[31,32,37,38])) or T_Timeout>5
              If AtHomePos or (In(ProgExe,[31,32,37,38]) and AtCenterPos)
                'nop'
              Else 
                Script: Report(90)
              If Progress_run() and  not ((digital_in[2] and ProgExe<50)  or (digital_in[6] and ProgExe>50))
                Script: Report(92)
            If Progress_run()
              Folder Camera
                MoveL speed 1000 mm/s, acceleration 3000 mm/s^2 (useActiveTCP=false optimoveEnabled=false optiMoveSpeed=0.3 optiMoveAcceleration=0.09) tcp=t0_Flange; feature=Base
                  If In(ProgExe,[31,32])
                    SetCameraProg := 32
                    Waypoint WpCenter: TCP in base x=62.197 y=393.251 z=616.502 mm, rx=-0.0356 ry=3.1413 rz=-0.0001 rad; joints [106.827, -57.183, -119.283, -93.604, 90.531, 15.582] deg; TCP offset x=0 y=0 z=0 mm, rx=0 ry=0 rz=3.1416 rad
                    Waypoint WLCamLMB: TCP in base x=6.314 y=481.622 z=313.228 mm, rx=0.3312 ry=3.1241 rz=0 rad; joints [110.281, -78.667, -139.534, -51.863, 90.366, 212.763] deg
                  If In(ProgExe,[37,38])
                    SetCameraProg := 37
                    Waypoint WpCenter: TCP in base x=62.197 y=393.251 z=616.502 mm, rx=-0.0356 ry=3.1413 rz=-0.0001 rad; joints [106.827, -57.183, -119.283, -93.604, 90.531, 15.582] deg; TCP offset x=0 y=0 z=0 mm, rx=0 ry=0 rz=3.1416 rad
                    Waypoint WLCamLMB2: TCP in base x=6.314 y=590.102 z=284.712 mm, rx=0.3312 ry=3.1241 rz=0 rad; joints [106.409, -92.678, -130.778, -46.608, 90.317, 28.92] deg
                  If In(ProgExe,[71,72])
                    SetCameraProg := 72
                    Waypoint WRBttnMidp: TCP in base x=1023.122 y=370.646 z=425.134 mm, rx=0 ry=3.1416 rz=0.0001 rad; joints [29.073, -130.015, -61.114, -78.934, 90.443, -60.761] deg; TCP offset x=0 y=0 z=0 mm, rx=0 ry=0 rz=3.1416 rad
                    Waypoint WRCamLMB: TCP in base x=1048.882 y=478.155 z=317.604 mm, rx=0.3312 ry=3.1241 rz=0 rad; joints [33.151, -139.694, -55, -75.371, 90.424, -44.561] deg; TCP offset x=0 y=0 z=0 mm, rx=0 ry=0 rz=3.1416 rad
                  If In(ProgExe,[77,78])
                    SetCameraProg := 77
                    Waypoint WRBttnMidp: TCP in base x=1023.122 y=370.646 z=425.134 mm, rx=0 ry=3.1416 rz=0.0001 rad; joints [29.073, -130.015, -61.114, -78.934, 90.443, -60.761] deg; TCP offset x=0 y=0 z=0 mm, rx=0 ry=0 rz=3.1416 rad
                    Waypoint WRCamLMB2: TCP in base x=1048.882 y=590.594 z=284.981 mm, rx=0.3312 ry=3.1241 rz=0 rad; joints [37.664, -146.75, -45.091, -78.225, 90.429, -40.076] deg; TCP offset x=0 y=0 z=0 mm, rx=0 ry=0 rz=3.1416 rad
                Call CamAcquire
                Call CamCalculateCorectnPlane
            If Progress_run() and CamCorrectnOK≠ProgExe
              MoveL speed 1000 mm/s, acceleration 3000 mm/s^2 (useActiveTCP=false optimoveEnabled=false optiMoveSpeed=0.3 optiMoveAcceleration=0.09) tcp=t0_Flange; feature=Base
                If ProgExe<50
                  Waypoint WpCenter: TCP in base x=62.197 y=393.251 z=616.502 mm, rx=-0.0356 ry=3.1413 rz=-0.0001 rad; joints [106.827, -57.183, -119.283, -93.604, 90.531, 15.582] deg
                  STS_Reservation := 0
                Else 
                  Waypoint WRBttnMidp: TCP in base x=1023.122 y=370.646 z=425.134 mm, rx=0 ry=3.1416 rz=0.0001 rad; joints [29.073, -130.015, -61.114, -78.934, 90.443, -60.761] deg; TCP offset x=0 y=0 z=0 mm, rx=0 ry=0 rz=3.1416 rad
                  Waypoint WRHome: TCP in base x=704.968 y=61.356 z=678.212 mm, rx=-2.2214 ry=-2.2214 rz=0 rad; joints [19.143, -89.513, -90.55, -90.002, 90.503, 19.233] deg; TCP offset x=0 y=0 z=0 mm, rx=0 ry=0 rz=3.1416 rad
              Script: Report(91)
            If Progress_run()
              Folder Lumbar
                If In(ProgExe,[31,32,37,38,71,72,77,78])
                  Timer (action=Reset) variable=T_Timeout
                  Timer (action=Start) variable=T_Timeout
                  Script: Report(12)
                  Wait Condition expression=Flags[2] or T_Timeout>60 or DEBUG or Abort
                  If Flags[2] or DEBUG
                    MoveL speed 1000 mm/s, acceleration 3000 mm/s^2 (useActiveTCP=false optimoveEnabled=false optiMoveSpeed=0.3 optiMoveAcceleration=0.09) tcp=t4_Finger; feature=Base
                      Folder Press FW
                        If False
                          Waypoint WLLmbFw: TCP in base x=-215.361 y=524.193 z=296.822 mm, rx=-0.3307 ry=-3.1201 rz=0.0016 rad; joints [113.232, -82.429, -130.104, -57.468, 90.623, 215.677] deg; TCP offset x=159 y=-58 z=70 mm, rx=0 ry=0 rz=0 rad
                          Waypoint WLLmbFw2: TCP in base x=-209.732 y=630.489 z=269.91 mm, rx=0.3312 ry=3.1241 rz=0 rad; joints [108.974, -94.642, -121.45, -53.973, 90.362, 31.442] deg; TCP offset x=-159 y=58 z=70 mm, rx=0 ry=0 rz=3.1416 rad
                          Waypoint WRLmbFw: TCP in base x=829.315 y=515.753 z=303.051 mm, rx=-0.3307 ry=-3.1201 rz=0.0016 rad; joints [37.179, -136.17, -55.721, -78.382, 90.551, 139.444] deg; TCP offset x=159 y=-58 z=70 mm, rx=0 ry=0 rz=0 rad
                          Waypoint WRLmbFw2: TCP in base x=826.645 y=629.264 z=271.348 mm, rx=0.3312 ry=3.1241 rz=0 rad; joints [41.665, -143.53, -45.442, -81.093, 90.438, -36.096] deg; TCP offset x=-159 y=58 z=70 mm, rx=0 ry=0 rz=3.1416 rad
                        If In(ProgExe,[31,32])
                          Wp := pose_add(WLLmbFw,Base_w_correctn)
                        If In(ProgExe,[37,38])
                          Wp := pose_add(WLLmbFw2,Base_w_correctn)
                        If In(ProgExe,[71,72])
                          Wp := pose_add(WRLmbFw,Base_w_correctn)
                        If In(ProgExe,[77,78])
                          Wp := pose_add(WRLmbFw2,Base_w_correctn)
                        Waypoint Variable (Variable): variable=Wp
                        Force Frame feature=Joint_6_name; selection=[1, 0, 0, 0, 0, 0]; wrench=[20, 10, -20, 0, 0, 0]; limitsForce=[0.05, 0.01, 0.05, 1.047198, 1.047198, 1.047198]; limitsMotion=[0.1, 0.1, 0.1, 0.349066, 0.349066, 0.349066]
                          Wait Sleep waitTime=0.7
                        ButtonPos := get_actual_tcp_pose()
                        Waypoint Variable (Variable): variable=Wp
                    Script: Report(3)
                  Else 
                    MoveL speed 1000 mm/s, acceleration 3000 mm/s^2 (useActiveTCP=false optimoveEnabled=false optiMoveSpeed=0.3 optiMoveAcceleration=0.09) tcp=t0_Flange; feature=Base
                      If ProgExe<50
                        Waypoint WpCenter: TCP in base x=62.197 y=393.251 z=616.502 mm, rx=-0.0356 ry=3.1413 rz=-0.0001 rad; joints [106.827, -57.183, -119.283, -93.604, 90.531, 15.582] deg; TCP offset x=0 y=0 z=0 mm, rx=0 ry=0 rz=3.1416 rad
                        STS_Reservation := 0
                      Else 
                        Waypoint WRBttnMidp: TCP in base x=1023.122 y=370.646 z=425.134 mm, rx=0 ry=3.1416 rz=0.0001 rad; joints [29.073, -130.015, -61.114, -78.934, 90.443, -60.761] deg; TCP offset x=0 y=0 z=0 mm, rx=0 ry=0 rz=3.1416 rad
                        Waypoint WRHome: TCP in base x=704.968 y=61.356 z=678.212 mm, rx=-2.2214 ry=-2.2214 rz=0 rad; joints [19.143, -89.513, -90.55, -90.002, 90.503, 19.233] deg; TCP offset x=0 y=0 z=0 mm, rx=0 ry=0 rz=3.1416 rad
                    Script: Report(95)
            If Progress_run()
              Folder Multiring
                If In(ProgExe,[32,38,72,78])
                  Timer (action=Reset) variable=T_Timeout
                  Timer (action=Start) variable=T_Timeout
                  Script: Report(11)
                  Wait Condition expression=Flags[1] or T_Timeout>60 or DEBUG or Abort
                  If Flags[1] or DEBUG
                    MoveL speed 1000 mm/s, acceleration 3000 mm/s^2 (useActiveTCP=false optimoveEnabled=false optiMoveSpeed=0.3 optiMoveAcceleration=0.09) tcp=t4_Finger; feature=Base
                      If False
                        Waypoint WLMultiringHi: TCP in base x=-236.485 y=507.422 z=309.965 mm, rx=0.2766 ry=3.1294 rz=0 rad; joints [116.04, -80.603, -129.951, -59.511, 90.408, 36.473] deg; TCP offset x=-159 y=58 z=70 mm, rx=0 ry=0 rz=3.1416 rad
                        Waypoint WLMultiringLo: TCP in base x=-234.901 y=510.523 z=286.198 mm, rx=-0.3307 ry=-3.1199 rz=0.0014 rad; joints [115.836, -81.881, -131.835, -56.263, 90.619, 218.29] deg; TCP offset x=159 y=-58 z=70 mm, rx=0 ry=0 rz=0 rad
                        Waypoint WLMultiringHi2: TCP in base x=-233.807 y=620.946 z=286.674 mm, rx=-0.3307 ry=-3.1199 rz=0.0014 rad; joints [111.267, -92.944, -121.349, -55.705, 90.611, 33.725] deg; TCP offset x=-159 y=58 z=70 mm, rx=0 ry=0 rz=3.1416 rad
                        Waypoint WLMultiringLo2: TCP in base x=-234.916 y=619.786 z=259.402 mm, rx=-0.3307 ry=-3.1199 rz=0.0014 rad; joints [111.399, -94.606, -122.911, -52.479, 90.59, 33.876] deg
                        Waypoint WRMultiringHi: TCP in base x=805.223 y=508.647 z=313.311 mm, rx=0.3312 ry=3.1241 rz=0 rad; joints [37.66, -133.152, -59.984, -76.93, 90.433, 139.942] deg; TCP offset x=159 y=-58 z=70 mm, rx=0 ry=0 rz=0 rad
                        Waypoint WRMultiringLo: TCP in base x=803.353 y=504.656 z=293.777 mm, rx=-0.3307 ry=-3.1199 rz=0.0014 rad; joints [37.531, -133.367, -61.653, -75.253, 90.557, 139.825] deg
                        Waypoint WRMultiringHi2: TCP in base x=805.086 y=620.683 z=282.502 mm, rx=0.3312 ry=3.1241 rz=0 rad; joints [42.055, -140.423, -50.073, -79.569, 90.436, -35.691] deg; TCP offset x=-159 y=58 z=70 mm, rx=0 ry=0 rz=3.1416 rad
                        Waypoint WRMultiringLo2: TCP in base x=805.256 y=618.494 z=260.601 mm, rx=0.3312 ry=3.1241 rz=0 rad; joints [41.966, -140.816, -51.588, -77.661, 90.43, -35.764] deg
                      Folder Press up
                        If ProgExe≟32
                          Wp0 := pose_add(WLMultiringLo,Base_w_correctn)
                        If ProgExe≟38
                          Wp0 := pose_add(WLMultiringLo2,Base_w_correctn)
                        If ProgExe≟72
                          Wp0 := pose_add(WRMultiringLo,Base_w_correctn)
                        If ProgExe≟78
                          Wp0 := pose_add(WRMultiringLo2,Base_w_correctn)
                        Wp0 := pose_trans(Wp0, p[-0.02,0,0,0,0,0])
                        Wp := Wp0
                        Script: Wp[0]=ButtonPos[0]-0.01
                        Waypoint Variable (Variable): variable=Wp0
                        Waypoint Variable (Variable): variable=Wp
                        Set NoAction tcp=t4_Finger
                        Force Frame feature=Joint_6_name; selection=[0, 1, 1, 0, 0, 0]; wrench=[10, 20, -20, 0, 0, 0]; limitsForce=[0.01, 0.01, 0.025, 1.047198, 1.047198, 1.047198]; limitsMotion=[0.1, 0.1, 0.1, 0.349066, 0.349066, 0.349066]
                          Wait Sleep waitTime=1
                        Waypoint Variable (Variable): variable=Wp0
                      Folder Press down
                        If ProgExe≟32
                          Wp0 := pose_add(WLMultiringHi,Base_w_correctn)
                        If ProgExe≟38
                          Wp0 := pose_add(WLMultiringHi2,Base_w_correctn)
                        If ProgExe≟72
                          Wp0 := pose_add(WRMultiringHi,Base_w_correctn)
                        If ProgExe≟78
                          Wp0 := pose_add(WRMultiringHi2,Base_w_correctn)
                        Wp0 := pose_trans(Wp0, p[-0.02,0,0,0,0,0])
                        Wp := Wp0
                        Script: Wp[0]=ButtonPos[0]-0.01
                        Waypoint Variable (Variable): variable=Wp0
                        Waypoint Variable (Variable): variable=Wp
                        Set NoAction tcp=t4_Finger
                        Force Frame feature=Joint_6_name; selection=[0, 1, 1, 0, 0, 0]; wrench=[10, 20, 20, 0, 0, 0]; limitsForce=[0.01, 0.01, 0.05, 1.047198, 1.047198, 1.047198]; limitsMotion=[0.1, 0.1, 0.1, 0.349066, 0.349066, 0.349066]
                          Wait Sleep waitTime=1
                        Waypoint Variable (Variable): variable=Wp0
                    Script: Report(2)
                  Else 
                    MoveL speed 1000 mm/s, acceleration 3000 mm/s^2 (useActiveTCP=false optimoveEnabled=false optiMoveSpeed=0.3 optiMoveAcceleration=0.09) tcp=t0_Flange; feature=Base
                      If ProgExe<50
                        Waypoint WpCenter: motionParameters(blendRadius=0.1); TCP in base x=62.197 y=393.251 z=616.502 mm, rx=-0.0356 ry=3.1413 rz=-0.0001 rad; joints [106.827, -57.183, -119.283, -93.604, 90.531, 15.582] deg; TCP offset x=0 y=0 z=0 mm, rx=0 ry=0 rz=3.1416 rad
                        STS_Reservation := 0
                      Else 
                        Waypoint WRBttnMidp: TCP in base x=1023.122 y=370.646 z=425.134 mm, rx=0 ry=3.1416 rz=0.0001 rad; joints [29.073, -130.015, -61.114, -78.934, 90.443, -60.761] deg; TCP offset x=0 y=0 z=0 mm, rx=0 ry=0 rz=3.1416 rad
                        Waypoint WRHome: TCP in base x=704.968 y=61.356 z=678.212 mm, rx=-2.2214 ry=-2.2214 rz=0 rad; joints [19.143, -89.513, -90.55, -90.002, 90.503, 19.233] deg; TCP offset x=0 y=0 z=0 mm, rx=0 ry=0 rz=3.1416 rad
                    Script: Report(95)
            If Progress_run()
              MoveL speed 1000 mm/s, acceleration 3000 mm/s^2 (useActiveTCP=false optimoveEnabled=false optiMoveSpeed=0.3 optiMoveAcceleration=0.09) tcp=t0_Flange; feature=Base
                If ProgExe<50
                  Waypoint WpCenter: TCP in base x=62.197 y=393.251 z=616.502 mm, rx=-0.0356 ry=3.1413 rz=-0.0001 rad; joints [106.827, -57.183, -119.283, -93.604, 90.531, 15.582] deg; TCP offset x=0 y=0 z=0 mm, rx=0 ry=0 rz=3.1416 rad
                  STS_Reservation := 0
                Else 
                  Waypoint WRBttnMidp: TCP in base x=1023.122 y=370.646 z=425.134 mm, rx=0 ry=3.1416 rz=0.0001 rad; joints [29.073, -130.015, -61.114, -78.934, 90.443, -60.761] deg; TCP offset x=0 y=0 z=0 mm, rx=0 ry=0 rz=3.1416 rad
                  Waypoint WRHome: TCP in base x=704.968 y=61.356 z=678.212 mm, rx=-2.2214 ry=-2.2214 rz=0 rad; joints [19.143, -89.513, -90.55, -90.002, 90.503, 19.233] deg; TCP offset x=0 y=0 z=0 mm, rx=0 ry=0 rz=3.1416 rad
              Script: Report(50)
        Folder Program finished
          ProgDn := ProgExe
          ProgExe := 0
      Folder Parking
        If Parking≟10 or ProgExe≟1010
          Wait Condition expression=EvtDock≤0
          If AtLHomePos
            MoveJ speed 120 deg/s, acceleration 500 deg/s^2 (useActiveTCP=true positionType=JointAngles optimoveEnabled=false optiMoveSpeed=0.3 optiMoveAcceleration=0.09) feature=Base
              Waypoint WpCenter: TCP in base x=62.197 y=393.251 z=616.502 mm, rx=-0.0356 ry=3.1413 rz=-0.0001 rad; joints [106.827, -57.183, -119.283, -93.604, 90.531, 15.582] deg; TCP offset x=0 y=0 z=0 mm, rx=0 ry=0 rz=3.1416 rad
          If AtRHomePos
            MoveJ speed 120 deg/s, acceleration 500 deg/s^2 (useActiveTCP=false positionType=JointAngles optimoveEnabled=false optiMoveSpeed=0.3 optiMoveAcceleration=0.09) tcp=t0_Flange; feature=Base
              Waypoint WRHome0: motionParameters(blendRadius=0.198); TCP in base x=228.171 y=378.753 z=507.074 mm, rx=1.3429 ry=2.8401 rz=-0.0001 rad; joints [62.572, -65.759, -114.23, -90.079, 90.522, 23.27] deg; TCP offset x=-134 y=56 z=118 mm, rx=0 ry=0 rz=3.1416 rad
              Waypoint WpCenter: TCP in base x=62.197 y=393.251 z=616.502 mm, rx=-0.0356 ry=3.1413 rz=-0.0001 rad; joints [106.827, -57.183, -119.283, -93.604, 90.531, 15.582] deg; TCP offset x=0 y=0 z=0 mm, rx=0 ry=0 rz=3.1416 rad
          Parking := 0
          If DEBUG
            ProgExe := 0
        If Parking≟11 or ProgExe≟1011
          Wait Condition expression=EvtDock≤0
          If AtLHomePos
            MoveJ speed 120 deg/s, acceleration 500 deg/s^2 (useActiveTCP=true positionType=JointAngles optimoveEnabled=false optiMoveSpeed=0.3 optiMoveAcceleration=0.09) feature=Base
              Waypoint WpCenter: motionParameters(blendRadius=0.1); TCP in base x=62.197 y=393.251 z=616.502 mm, rx=-0.0356 ry=3.1413 rz=-0.0001 rad; joints [106.827, -57.183, -119.283, -93.604, 90.531, 15.582] deg
              Waypoint WpParkUp0: motionParameters(blendRadius=0.1); TCP in base x=174.17 y=174.659 z=748.205 mm, rx=-2.2127 ry=2.2111 rz=0.001 rad; joints [90.202, -42.467, -109.682, -117.347, 90, -89.999] deg
              Waypoint WpPark: TCP in base x=175.046 y=118.455 z=1248.983 mm, rx=-2.2111 ry=2.2293 rz=-0.0002 rad; joints [89.999, -90, 0, -180, 90, -90] deg
          If AtRHomePos
            MoveJ speed 120 deg/s, acceleration 500 deg/s^2 (useActiveTCP=false positionType=JointAngles optimoveEnabled=false optiMoveSpeed=0.3 optiMoveAcceleration=0.09) tcp=t0_Flange; feature=Base
              Waypoint WRHome0: motionParameters(blendRadius=0.2); TCP in base x=228.171 y=378.753 z=507.074 mm, rx=1.3429 ry=2.8401 rz=-0.0001 rad; joints [62.572, -65.759, -114.23, -90.079, 90.522, 23.27] deg; TCP offset x=-134 y=56 z=118 mm, rx=0 ry=0 rz=3.1416 rad
              Waypoint WpCenter: motionParameters(blendRadius=0.1); TCP in base x=62.197 y=393.251 z=616.502 mm, rx=-0.0356 ry=3.1413 rz=-0.0001 rad; joints [106.827, -57.183, -119.283, -93.604, 90.531, 15.582] deg; TCP offset x=0 y=0 z=0 mm, rx=0 ry=0 rz=3.1416 rad
              Waypoint WpParkUp0: motionParameters(blendRadius=0.1); TCP in base x=174.17 y=174.659 z=748.205 mm, rx=-2.2127 ry=2.2111 rz=0.001 rad; joints [90.202, -42.467, -109.682, -117.347, 90, -89.999] deg
              Waypoint WpPark: TCP in base x=175.046 y=118.455 z=1248.983 mm, rx=-2.2111 ry=2.2293 rz=-0.0002 rad; joints [89.999, -90, 0, -180, 90, -90] deg
              SuppressedNode
                Waypoint WpParkOld: TCP in base x=53.158 y=791.824 z=735.444 mm, rx=-0.0355 ry=3.1413 rz=-0.0001 rad; joints [98.778, -98.151, -75.54, -96.378, 90.491, 7.516] deg
          If AtCenterPos
            MoveJ speed 120 deg/s, acceleration 500 deg/s^2 (useActiveTCP=false positionType=JointAngles optimoveEnabled=false optiMoveSpeed=0.3 optiMoveAcceleration=0.09) tcp=t0_Flange; feature=Base
              Waypoint WpParkUp0: motionParameters(blendRadius=0.1); TCP in base x=174.17 y=174.659 z=748.205 mm, rx=-2.2127 ry=2.2111 rz=0.001 rad; joints [90.202, -42.467, -109.682, -117.347, 90, -89.999] deg
              Waypoint WpPark: TCP in base x=175.046 y=118.455 z=1248.983 mm, rx=-2.2111 ry=2.2293 rz=-0.0002 rad; joints [89.999, -90, 0, -180, 90, -90] deg
          Parking := 0
          If DEBUG
            ProgExe := 0
        If Parking≟1 or ProgExe≟1001
          If AtParkPos
            MoveJ speed 120 deg/s, acceleration 500 deg/s^2 (useActiveTCP=false positionType=JointAngles optimoveEnabled=false optiMoveSpeed=0.3 optiMoveAcceleration=0.09) tcp=t0_Flange; feature=Base
              Waypoint WpParkUp0: motionParameters(blendRadius=0.1); TCP in base x=174.17 y=174.659 z=748.205 mm, rx=-2.2127 ry=2.2111 rz=0.001 rad; joints [90.202, -42.467, -109.682, -117.347, 90, -89.999] deg
              Waypoint WpCenter: motionParameters(blendRadius=0.1); TCP in base x=62.197 y=393.251 z=616.502 mm, rx=-0.0356 ry=3.1413 rz=-0.0001 rad; joints [106.827, -57.183, -119.283, -93.604, 90.531, 15.582] deg
              Waypoint WLHome: TCP in base x=-773.534 y=70.689 z=655.308 mm, rx=3.1416 ry=0 rz=0 rad; joints [187.663, -96.209, -85.791, -88.066, 90.49, -82.232] deg
              STS_Reservation := 1
          If AtCenterPos
            MoveJ speed 120 deg/s, acceleration 500 deg/s^2 (useActiveTCP=false positionType=JointAngles optimoveEnabled=false optiMoveSpeed=0.3 optiMoveAcceleration=0.09) tcp=t0_Flange; feature=Base
              Waypoint WLHome: TCP in base x=-773.534 y=70.689 z=655.308 mm, rx=3.1416 ry=0 rz=0 rad; joints [187.663, -96.209, -85.791, -88.066, 90.49, -82.232] deg
              STS_Reservation := 1
          If AtRHomePos
            MoveJ speed 120 deg/s, acceleration 500 deg/s^2 (useActiveTCP=false positionType=JointAngles optimoveEnabled=false optiMoveSpeed=0.3 optiMoveAcceleration=0.09) tcp=t0_Flange; feature=Base
              Waypoint WRHome0: motionParameters(blendRadius=0.107); TCP in base x=228.171 y=378.753 z=507.074 mm, rx=1.3429 ry=2.8401 rz=-0.0001 rad; joints [62.572, -65.759, -114.23, -90.079, 90.522, 23.27] deg; TCP offset x=-134 y=56 z=118 mm, rx=0 ry=0 rz=3.1416 rad
              Waypoint WpCenter: motionParameters(blendRadius=0.091); TCP in base x=62.197 y=393.251 z=616.502 mm, rx=-0.0356 ry=3.1413 rz=-0.0001 rad; joints [106.827, -57.183, -119.283, -93.604, 90.531, 15.582] deg; TCP offset x=0 y=0 z=0 mm, rx=0 ry=0 rz=3.1416 rad
              Waypoint WLHome: TCP in base x=-773.534 y=70.689 z=655.308 mm, rx=3.1416 ry=0 rz=0 rad; joints [187.663, -96.209, -85.791, -88.066, 90.49, -82.232] deg
              STS_Reservation := 1
          Parking := 0
          If DEBUG
            ProgExe := 0
        If Parking≟2 or ProgExe≟1002
          If AtParkPos
            MoveJ speed 120 deg/s, acceleration 500 deg/s^2 (useActiveTCP=false positionType=JointAngles optimoveEnabled=false optiMoveSpeed=0.3 optiMoveAcceleration=0.09) tcp=t0_Flange; feature=Base
              Waypoint WpParkUp0: motionParameters(blendRadius=0.1); TCP in base x=174.17 y=174.659 z=748.205 mm, rx=-2.2127 ry=2.2111 rz=0.001 rad; joints [90.202, -42.467, -109.682, -117.347, 90, -89.999] deg
              Waypoint WpCenter: motionParameters(blendRadius=0.091); TCP in base x=62.197 y=393.251 z=616.502 mm, rx=-0.0356 ry=3.1413 rz=-0.0001 rad; joints [106.827, -57.183, -119.283, -93.604, 90.531, 15.582] deg
              Waypoint WRHome0: motionParameters(blendRadius=0.2); TCP in base x=228.171 y=378.753 z=507.074 mm, rx=1.3429 ry=2.8401 rz=-0.0001 rad; joints [62.572, -65.759, -114.23, -90.079, 90.522, 23.27] deg; TCP offset x=-134 y=56 z=118 mm, rx=0 ry=0 rz=3.1416 rad
              Waypoint WRHome: TCP in base x=704.968 y=61.356 z=678.212 mm, rx=-2.2214 ry=-2.2214 rz=0 rad; joints [19.143, -89.513, -90.55, -90.002, 90.503, 19.233] deg; TCP offset x=0 y=0 z=0 mm, rx=0 ry=0 rz=3.1416 rad
              STS_Reservation := 2
          If AtCenterPos
            MoveJ speed 120 deg/s, acceleration 500 deg/s^2 (useActiveTCP=true positionType=JointAngles optimoveEnabled=false optiMoveSpeed=0.3 optiMoveAcceleration=0.09) feature=Base
              Waypoint WRHome0: motionParameters(blendRadius=0.198); TCP in base x=228.171 y=378.753 z=507.074 mm, rx=1.3429 ry=2.8401 rz=-0.0001 rad; joints [62.572, -65.759, -114.23, -90.079, 90.522, 23.27] deg; TCP offset x=-134 y=56 z=118 mm, rx=0 ry=0 rz=3.1416 rad
              Waypoint WRHome: TCP in base x=704.968 y=61.356 z=678.212 mm, rx=-2.2214 ry=-2.2214 rz=0 rad; joints [19.143, -89.513, -90.55, -90.002, 90.503, 19.233] deg; TCP offset x=0 y=0 z=0 mm, rx=0 ry=0 rz=3.1416 rad
              STS_Reservation := 2
          If AtLHomePos
            MoveJ speed 120 deg/s, acceleration 500 deg/s^2 (useActiveTCP=false positionType=JointAngles optimoveEnabled=false optiMoveSpeed=0.3 optiMoveAcceleration=0.09) tcp=t0_Flange; feature=Base
              Waypoint WpCenter: motionParameters(blendRadius=0.048); TCP in base x=62.197 y=393.251 z=616.502 mm, rx=-0.0356 ry=3.1413 rz=-0.0001 rad; joints [106.827, -57.183, -119.283, -93.604, 90.531, 15.582] deg; TCP offset x=0 y=0 z=0 mm, rx=0 ry=0 rz=3.1416 rad
              Waypoint WRHome0: motionParameters(blendRadius=0.15); TCP in base x=228.171 y=378.753 z=507.074 mm, rx=1.3429 ry=2.8401 rz=-0.0001 rad; joints [62.572, -65.759, -114.23, -90.079, 90.522, 23.27] deg; TCP offset x=-134 y=56 z=118 mm, rx=0 ry=0 rz=3.1416 rad
              Waypoint WRHome: TCP in base x=704.968 y=61.356 z=678.212 mm, rx=-2.2214 ry=-2.2214 rz=0 rad; joints [19.143, -89.513, -90.55, -90.002, 90.503, 19.233] deg; TCP offset x=0 y=0 z=0 mm, rx=0 ry=0 rz=3.1416 rad
              STS_Reservation := 2
          Parking := 0
          If DEBUG
            ProgExe := 0
Thread Thread_1 (runOnlyOnce=false)
  Folder Continuous calculations
    Folder get live force and tcp pos
      P_act := get_actual_tcp_pose()
      V_act := get_actual_tcp_speed()
      V_act_norm := norm(V_act)
      P_Flange := get_actual_tool_flange_pose()
      D_rel := pose_sub(P_act, P_ini)
      Folder Detect home positions
        AtLHomePos := PosDist(P_Flange, WLHome)<0.005
        AtRHomePos := PosDist(P_Flange, WRHome)<0.005
        AtCenterPos := PosDist(P_Flange, WpCenter)<0.005
        AtParkPos := PosDist(P_Flange, WpPark)<0.005
        If InRange(ProgExe,10,49)
          AtHomePos := AtLHomePos
        ElseIf InRange(ProgExe,50,89)
          AtHomePos := AtRHomePos
        Else 
          AtHomePos := AtLHomePos or AtRHomePos
      Folder Detect docking signal
        If P_Flange[0]<0
          AdapterDocked := digital_in[0]
        Else 
          AdapterDocked := digital_in[4]
      Folder Calculate actual offset in tool frame
        If ProgExe≟15
          TempWp := pose_sub(WLBuckleSpa1,Base_w_correctn)
          BklToolDist := pose_trans(pose_inv(TempWp), P_act)
        If ProgExe≟16
          TempWp := pose_sub(WLBuckleSpa3,Base_w_correctn)
          BklToolDist := pose_trans(pose_inv(TempWp), P_act)
        If ProgExe≟55
          TempWp := pose_sub(WRBuckleSpa1,Base_w_correctn)
          BklToolDist := pose_trans(pose_inv(TempWp), P_act)
        If ProgExe≟56
          TempWp := pose_sub(WRBuckleSpa3,Base_w_correctn)
          BklToolDist := pose_trans(pose_inv(TempWp), P_act)
      Folder InterlockOutput
        If P_Flange[1]<0.45
          Set DigitalOutput pin=digital_out[7]; digitalValue=1
        ElseIf P_Flange[0]>0.65
          Set DigitalOutput pin=digital_out[7]; digitalValue=1
        ElseIf InRange(P_Flange[0],-0.35,0)
          Set DigitalOutput pin=digital_out[7]; digitalValue=1
        Else 
          Set DigitalOutput pin=digital_out[7]; digitalValue=0
    Folder Modbus mapping
      Folder Heartbeat
        Timer (action=Start) variable(name=T_Heartbeat)
        If T_Heartbeat≥1
          Timer (action=Reset) variable=T_Heartbeat
          If STS_Heartbeat
            STS_Heartbeat := False
          Else 
            STS_Heartbeat := True
      Folder Safe position
        Folder L
          STS_Safe_i1 := True
          If pose_dist(P_act, WLConnSpa1)<0.08
            STS_Safe_i1 := False
          If pose_dist(P_act, WLUnplug1_3)<0.05
            STS_Safe_i1 := False
          If pose_dist(P_act, WLBuckleSpa1)<0.2
            STS_Safe_i1 := False
          If pose_dist(P_act, WLLmbFw)<0.05
            STS_Safe_i1 := False
          If pose_dist(P_act, WLLmbFw2)<0.05
            STS_Safe_i1 := False
        Folder R
          STS_Safe_i2 := True
          If pose_dist(P_act, WRConnSpa1)<0.08
            STS_Safe_i2 := False
          If pose_dist(P_act, WRUnpgSpa1_4)<0.05
            STS_Safe_i2 := False
          If pose_dist(P_act, WRBuckleSpa1)<0.2
            STS_Safe_i2 := False
          If pose_dist(P_act, WRLmbFw)<0.05
            STS_Safe_i2 := False
          If pose_dist(P_act, WRLmbFw2)<0.05
            STS_Safe_i2 := False
      Folder Outputs
        Script: write_port_register(129,STS_Progress)
        Script: write_port_register(131,STS_Reservation)
        Script: write_port_register(134,binary_list_to_integer([digital_in[0],digital_in[4],config_in[0],STS_Heartbeat,STS_Safe_i1,STS_Safe_i2]))
      Folder Inputs
        CMD_Reserve_i1 := read_port_register(160)
        CMD_Reserve_i2 := read_port_register(161)
        CMD_Timeout_i1 := read_port_register(162)
        CMD_Timeout_i2 := read_port_register(163)
        CMD_Program_i1 := read_port_register(164)
        CMD_Program_i2 := read_port_register(165)
        CMD_Flags_i1 := read_port_register(170)
        CMD_Flags_i2 := read_port_register(171)
        CMD_Heartbt_i1 := read_port_register(180)
        CMD_Heartbt_i2 := read_port_register(181)
      Folder Generate flags
        Flags_i1 := integer_to_binary_list(CMD_Flags_i1)
        Flags_i2 := integer_to_binary_list(CMD_Flags_i2)
        If InRange(ProgExe,10,49)
          Flags := Flags_i1
        ElseIf InRange(ProgExe,50,89)
          Flags := Flags_i2
    Folder Operator call deactivation
      If digital_out[1] or digital_out[2]
        Timer (action=Start) variable(name=T_Call)
        If not  NormalMode and T_Call>4
          Set DigitalOutput pin=digital_out[1]; digitalValue=0
          Set DigitalOutput pin=digital_out[2]; digitalValue=0
          Mute := True
      Else 
        Timer (action=Stop) variable=T_Call
        Timer (action=Reset) variable=T_Call
      If ProgExe>0
        Mute := False
    Folder Abort
      If Flags_i1[14] and (InRange(ProgExe,10,49) or AdapterReady_L)
        Abort := True
      ElseIf Flags_i2[14] and (InRange(ProgExe,50,89) or AdapterReady_R)
        Abort := True
      If AtHomePos or AtCenterPos
        Abort := False
      If Abort
        If AdapterReady_L or AdapterReady_R
          EvtDock := 1
    Folder Speed
      Timer (action=Start) variable(name=T_SpeedSet)
      If T_SpeedSet>2 and  not DEBUG
        Script: socket_send_string("set speed")
        Script: socket_send_string(1.0)
        Script: socket_send_byte(10)
        Timer (action=Reset) variable=T_SpeedSet
    Wait Sleep waitTime=0.01
  Folder ReservationControl
    'Request reservation, disconnect preference'
    If STS_Reservation≟0 and ProgExe≟0 and Parking≟0
      If CMD_Reserve_i1≟1 and In(CMD_Program_i1,[21,22,23])
        'request reservation'
        If AtLHomePos or AdapterReady_L
          STS_Reservation := 1
        Else 
          Parking := 1
      If CMD_Reserve_i2≟2 and In(CMD_Program_i2,[61,62,63])
        'request reservation'
        If AtRHomePos or AdapterReady_R
          STS_Reservation := 2
        Else 
          Parking := 2
      If CMD_Reserve_i1≟1
        'request reservation'
        If AtLHomePos or AdapterReady_L
          STS_Reservation := 1
        ElseIf In(CMD_Program_i1,[31,32,37,38])
          'Special case to save time when moving to buttons'
          If AtCenterPos
            STS_Reservation := 1
          Else 
            Parking := 10
        Else 
          Parking := 1
      If CMD_Reserve_i2≟2
        'request reservation'
        If AtRHomePos or AdapterReady_R
          STS_Reservation := 2
        ElseIf In(CMD_Program_i2,[55,56])
          'Special case to save time when moving to buckle'
          If AtCenterPos
            STS_Reservation := 2
          Else 
            Parking := 10
        Else 
          Parking := 2
    'Timeout reservation - station keeps reservation for a while to prevent other app stealing the process'
    'Timeout is configurable, so application can control how long to keep robot before letting other app'
    If STS_Progress≟0 and STS_Reservation≠0 and Parking≟0
      If STS_Reservation≟1 and CMD_Reserve_i1≟1
        'nop'
      ElseIf STS_Reservation≟2 and CMD_Reserve_i2≟2
        'nop'
      Else 
        If STS_Reservation≟1
          T_KeepReservtn := CMD_Timeout_i1
        If STS_Reservation≟2
          T_KeepReservtn := CMD_Timeout_i2
        Timer (action=Start) variable(name=T_Unreserve)
        If T_Unreserve>T_KeepReservtn
          STS_Reservation := 0
    Else 
      Timer (action=Stop) variable=T_Unreserve
      Timer (action=Reset) variable=T_Unreserve
    'Force release reservation from app - in case of intervetion'
    If STS_Reservation≟0 and STS_Progress≟0 and  not DEBUG
      If In(CMD_Reserve_i1,[98,99]) and  not In(CMD_Reserve_i2,[98,99]) and  not AtParkPos
        If AtRHomePos
          STS_Reservation := 2
        Else 
          Parking := 2
      If In(CMD_Reserve_i2,[98,99]) and  not In(CMD_Reserve_i1,[98,99]) and  not AtParkPos
        If AtLHomePos
          STS_Reservation := 1
        Else 
          Parking := 1
      If In(CMD_Reserve_i1,[98,99]) and In(CMD_Reserve_i2,[98,99])
        If AtParkPos
          STS_Reservation := 0
        Else 
          Parking := 11
      If (CMD_Reserve_i1≟99 or CMD_Reserve_i2≟99) and  not Mute
        Set DigitalOutput pin=digital_out[1]; digitalValue=1
        Set DigitalOutput pin=digital_out[2]; digitalValue=1
  Folder Program control
    'Start new Prog / Confirm Prog Running'
    If STS_Progress≟0 and ProgExe≟0  and  not Abort and  not DEBUG
      If InRange(CMD_Program_i1,10,49) and STS_Reservation≟1
        ProgExe := CMD_Program_i1
        T_KeepReservtn := CMD_Timeout_i1
        Script: Report(0)
      If InRange(CMD_Program_i2,50,89) and STS_Reservation≟2
        ProgExe := CMD_Program_i2
        T_KeepReservtn := CMD_Timeout_i2
        Script: Report(0)
    'Ack results - get ready for new prg'
    If ProgExe≟0 and Progress_finished()
      If InRange(ProgDn,10,49) and CMD_Program_i1≠ProgDn
        STS_Progress := 0
        If In(CMD_Program_i1,[21,22,23]) or In(CMD_Program_i2,[61,62,63])
          'unplug preference - unreserve immediatelly'
          STS_Reservation := 0
      If InRange(ProgDn,50,89) and CMD_Program_i2≠ProgDn
        STS_Progress := 0
        If In(CMD_Program_i1,[21,22,23]) or In(CMD_Program_i2,[61,62,63])
          'unplug preference - unreserve immediatelly'
          STS_Reservation := 0
SubProgram WaitForNormalMode [hidden by the author, left out]
SubProgram  [hidden by the author, left out]
SubProgram  [hidden by the author, left out]
SubProgram  [hidden by the author, left out]
SubProgram  [hidden by the author, left out]
Event  expression=SetCameraProg>0
  Folder Set program to camera in advance
    Set DigitalOutput pin=CnxDO_Trig; digitalValue=0
    Set DigitalOutput pin=CnxDO_TrigEn; digitalValue=1
    Script: modbus_delete_signal("CnxAO_Program")
    Script: modbus_add_signal("10.142.142.41", 255, 2001, 16, "CnxAO_Program", True ,1)
    Script: modbus_set_output_register("CnxAO_Program",SetCameraProg, False )
    Wait Sleep waitTime=0.2
    Set DigitalOutput pin=CnxDO_SetUsrDta; digitalValue=1
    Wait DigitalInput pin=CnxDi_UsrDtaAck; digitalValue=1
    Set DigitalOutput pin=CnxDO_SetUsrDta; digitalValue=0
    Set DigitalOutput pin=CnxDO_SoftEvt0; digitalValue=1
    Wait DigitalInput pin=CnxDI_Evt0Ack; digitalValue=1
    Set DigitalOutput pin=CnxDO_SoftEvt0; digitalValue=0
    Timer (action=Reset) variable=CamTimeout
    Timer (action=Start) variable=CamTimeout
    Wait Condition expression=CnxAI_Program≟SetCameraProg or CamTimeout>3
    If CnxAI_Program≠SetCameraProg
      Script: textmsg("set cam prog failed, trying trigger")
      Folder For the first time it needs trigger when going online
        Set DigitalOutput pin=CnxDO_Trig; digitalValue=1
        Wait Sleep waitTime=1
        Set DigitalOutput pin=CnxDO_Trig; digitalValue=0
      If CnxAI_Program≠SetCameraProg
        SuppressedNode
          Popup Error (haltProgram=false message=Error: camera program not set inputType=Text)
      Else 
        Wait Sleep waitTime=0.5
        SetCameraProg := 0
    Else 
      Wait Sleep waitTime=0.5
      SetCameraProg := 0
  If SetCameraProg>0
    'repeat on fail'
    Wait Sleep waitTime=3
    Folder Set program to camera in advance
      Set DigitalOutput pin=CnxDO_Trig; digitalValue=0
      Set DigitalOutput pin=CnxDO_TrigEn; digitalValue=1
      Script: modbus_delete_signal("CnxAO_Program")
      Script: modbus_add_signal("10.142.142.41", 255, 2001, 16, "CnxAO_Program", True ,1)
      Script: modbus_set_output_register("CnxAO_Program",SetCameraProg, False )
      Wait Sleep waitTime=0.2
      Set DigitalOutput pin=CnxDO_SetUsrDta; digitalValue=1
      Wait DigitalInput pin=CnxDi_UsrDtaAck; digitalValue=1
      Set DigitalOutput pin=CnxDO_SetUsrDta; digitalValue=0
      Set DigitalOutput pin=CnxDO_SoftEvt0; digitalValue=1
      Wait DigitalInput pin=CnxDI_Evt0Ack; digitalValue=1
      Set DigitalOutput pin=CnxDO_SoftEvt0; digitalValue=0
      Timer (action=Reset) variable=CamTimeout
      Timer (action=Start) variable=CamTimeout
      Wait Condition expression=CnxAI_Program≟SetCameraProg or CamTimeout>3
      If CnxAI_Program≠SetCameraProg
        Script: textmsg("set cam prog failed, trying trigger")
        Folder For the first time it needs trigger when going online
          Set DigitalOutput pin=CnxDO_Trig; digitalValue=1
          Wait Sleep waitTime=1
          Set DigitalOutput pin=CnxDO_Trig; digitalValue=0
        If CnxAI_Program≠SetCameraProg
          SuppressedNode
            Popup Error (haltProgram=false message=Error: camera program not set inputType=Text)
        Else 
          Wait Sleep waitTime=0.5
          SetCameraProg := 0
      Else 
        Wait Sleep waitTime=0.5
        SetCameraProg := 0
  If SetCameraProg>0
    'repeat on fail'
    Wait Sleep waitTime=3
    Folder Set program to camera in advance
      Set DigitalOutput pin=CnxDO_Trig; digitalValue=0
      Set DigitalOutput pin=CnxDO_TrigEn; digitalValue=1
      Script: modbus_delete_signal("CnxAO_Program")
      Script: modbus_add_signal("10.142.142.41", 255, 2001, 16, "CnxAO_Program", True ,1)
      Script: modbus_set_output_register("CnxAO_Program",SetCameraProg, False )
      Wait Sleep waitTime=0.2
      Set DigitalOutput pin=CnxDO_SetUsrDta; digitalValue=1
      Wait DigitalInput pin=CnxDi_UsrDtaAck; digitalValue=1
      Set DigitalOutput pin=CnxDO_SetUsrDta; digitalValue=0
      Set DigitalOutput pin=CnxDO_SoftEvt0; digitalValue=1
      Wait DigitalInput pin=CnxDI_Evt0Ack; digitalValue=1
      Set DigitalOutput pin=CnxDO_SoftEvt0; digitalValue=0
      Timer (action=Reset) variable=CamTimeout
      Timer (action=Start) variable=CamTimeout
      Wait Condition expression=CnxAI_Program≟SetCameraProg or CamTimeout>3
      If CnxAI_Program≠SetCameraProg
        Script: textmsg("set cam prog failed, trying trigger")
        Folder For the first time it needs trigger when going online
          Set DigitalOutput pin=CnxDO_Trig; digitalValue=1
          Wait Sleep waitTime=1
          Set DigitalOutput pin=CnxDO_Trig; digitalValue=0
        If CnxAI_Program≠SetCameraProg
          SuppressedNode
            Popup Error (haltProgram=false message=Error: camera program not set inputType=Text)
        Else 
          Wait Sleep waitTime=0.5
          SetCameraProg := 0
      Else 
        Wait Sleep waitTime=0.5
        SetCameraProg := 0
  If SetCameraProg>0
    Popup Error (haltProgram=false message=Error: camera program not set inputType=Text)
SubProgram -> CamAcquire
SubProgram -> CamCalculateCorectnPlane
Event  expression=EvtDock>0
  Folder Dock
    MoveL speed 1000 mm/s, acceleration 3000 mm/s^2 (useActiveTCP=false optimoveEnabled=false optiMoveSpeed=0.3 optiMoveAcceleration=0.09) tcp=t2_Gripper; feature=Base
      If EvtDock≟2
        Folder Force mvts
          Set NoAction tcp=t2_Gripper
          Wp0 := P_act
          Force Frame feature=Joint_6_name; selection=[0, 1, 0, 0, 0, 0]; wrench=[0, -20, 0, 0, 0, 0]; limitsForce=[0.15, 0.1, 0.15, 1.047198, 1.047198, 1.047198]; limitsMotion=[0.1, 0.1, 0.1, 0.349066, 0.349066, 0.349066]
            Wait Sleep waitTime=1
          Force Frame feature=Joint_6_name; selection=[1, 0, 1, 1, 0, 0]; wrench=[0, -10, 0, 0, 0, 0]; limitsForce=[0.15, 0.05, 0.1, 1.047198, 1.047198, 1.047198]; limitsMotion=[0.1, 0.1, 0.1, 0.349066, 0.349066, 0.349066]
            Wait Sleep waitTime=0.2
            Call GripperClose
            Wait Sleep waitTime=0.2
          If T_Gripper>3
            Call GripperOpen
            MoveL speed 500 mm/s, acceleration 1200 mm/s^2 (useActiveTCP=true optimoveEnabled=false optiMoveSpeed=0.3 optiMoveAcceleration=0.09) feature=Base
              Waypoint Variable (Variable): variable=Wp0
            Force Frame feature=Joint_6_name; selection=[0, 1, 0, 0, 0, 0]; wrench=[0, -20, 0, 0, 0, 0]; limitsForce=[0.15, 0.1, 0.15, 1.047198, 1.047198, 1.047198]; limitsMotion=[0.1, 0.1, 0.1, 0.349066, 0.349066, 0.349066]
              Wait Sleep waitTime=1
            Force Frame feature=Joint_6_name; selection=[1, 0, 1, 0, 0, 0]; wrench=[0, -10, 0, 0, 0, 0]; limitsForce=[0.15, 0.05, 0.1, 1.047198, 1.047198, 1.047198]; limitsMotion=[0.1, 0.1, 0.1, 0.349066, 0.349066, 0.349066]
              Wait Sleep waitTime=0.2
              Call GripperClose
              Wait Sleep waitTime=0.2
          If T_Gripper>3
            Call GripperOpen
            MoveL speed 500 mm/s, acceleration 1200 mm/s^2 (useActiveTCP=true optimoveEnabled=false optiMoveSpeed=0.3 optiMoveAcceleration=0.09) feature=Base
              Waypoint Variable (Variable): variable=Wp0
              EvtDock := -97
          If EvtDock≟2
            MoveDirectionNode (selectedDirection=YPlus) feature=Joint_6_name
              Until DISTANCE (allowActions=false deceleration=3 distanceNodeType=BLEND) Distance=0.1; motionParameters(blendRadius=0.05)
      If InRange(EvtDock,1,2)
        If P_Flange[0]<0
          WpDock := WLDock
          WpHome := WLHome
        Else 
          WpDock := WRDock
          WpHome := WRHome
        Script: Report(40)
        Wp := pose_trans(WpDock, p[0,0.25,0,0,0,0])
        Waypoint Variable (Variable): motionParameters(blendRadius=0.05); variable=Wp
        Waypoint Variable (Variable): variable=WpDock
        Call GripperOpen
        Waypoint Variable (Variable): variable=Wp
        MoveL speed 1000 mm/s, acceleration 3000 mm/s^2 (useActiveTCP=false optimoveEnabled=false optiMoveSpeed=0.3 optiMoveAcceleration=0.09) tcp=t0_Flange; feature=Base
          Waypoint Variable (Variable): variable=WpHome
        EvtDock := 0
Event  expression=EvtBeep
  Loop While (checkContinuously=false) expression=EvtBeep
    Set DigitalOutput pin=digital_out[2]; digitalValue=1
    Set DigitalOutput pin=digital_out[1]; digitalValue=1
    Wait Sleep waitTime=0.5
    Set DigitalOutput pin=digital_out[2]; digitalValue=0
    Set DigitalOutput pin=digital_out[1]; digitalValue=0
    Wait Sleep waitTime=5
SubProgram GripperOpen [hidden by the author, left out]
SubProgram GripperOpenQuick [hidden by the author, left out]
SubProgram GripperClose [hidden by the author, left out]
SubProgram CamAcquire (keepSynchronizedWithDisk=false)
  Folder Trig camera and process data
    Folder Init
      CamCorrectnOK := 0
      CamRetry := 0
    Wait Condition expression=SetCameraProg≟0
    Loop While (checkContinuously=false) expression=CamRetry<3
      Folder Trig
        CnxCounter := CnxAI_Counter
        Set DigitalOutput pin=CnxDO_Trig; digitalValue=1
        Timer (action=Reset) variable(name=CamTimeout)
        Timer (action=Start) variable=CamTimeout
        Wait Condition expression=CamTimeout>1 or CnxAI_Counter≠CnxCounter
        Set DigitalOutput pin=CnxDO_Trig; digitalValue=0
        Wait Sleep waitTime=0.2
        If CnxAI_Result≥100 and CnxAI_Counter≠CnxCounter
          CamRetry := 100
        Else 
          Wait Sleep waitTime=1
          CamRetry := CamRetry+1
    Folder New data validation
      If CamRetry≟100
        CamCorrectnOK := ProgExe
      Else 
        CamCorrectnOK := 0
      CamData := [(CnxAI_ResultX-30000)/10000,(CnxAI_ResultY-30000)/10000,d2r((CnxAI_ResultR-30000)/10)]
      SuppressedNode
        If CamData[1]>0.03
          Err_state := 103
      SuppressedNode
        If CamData[1]<-0.03
          Err_state := 104
      SuppressedNode
        If CamData[2]>15
          Err_state := 105
      SuppressedNode
        If CamData[2]<-15
          Err_state := 106
SubProgram GripperCloseQuick [hidden by the author, left out]
SubProgram CamCalculateCorectnPlane (keepSynchronizedWithDisk=false)
  Folder Folder
    Set NoAction tcp=t0_Flange
    Script: sync()
    P_act := get_actual_tcp_pose()
    CamCorrection := p[0,CamData[0],CamData[1],0,0,0]
    CamOffset := pose_trans(P_act,CamCorrection)
    Base_w_correctn := pose_sub(CamOffset, P_act)
